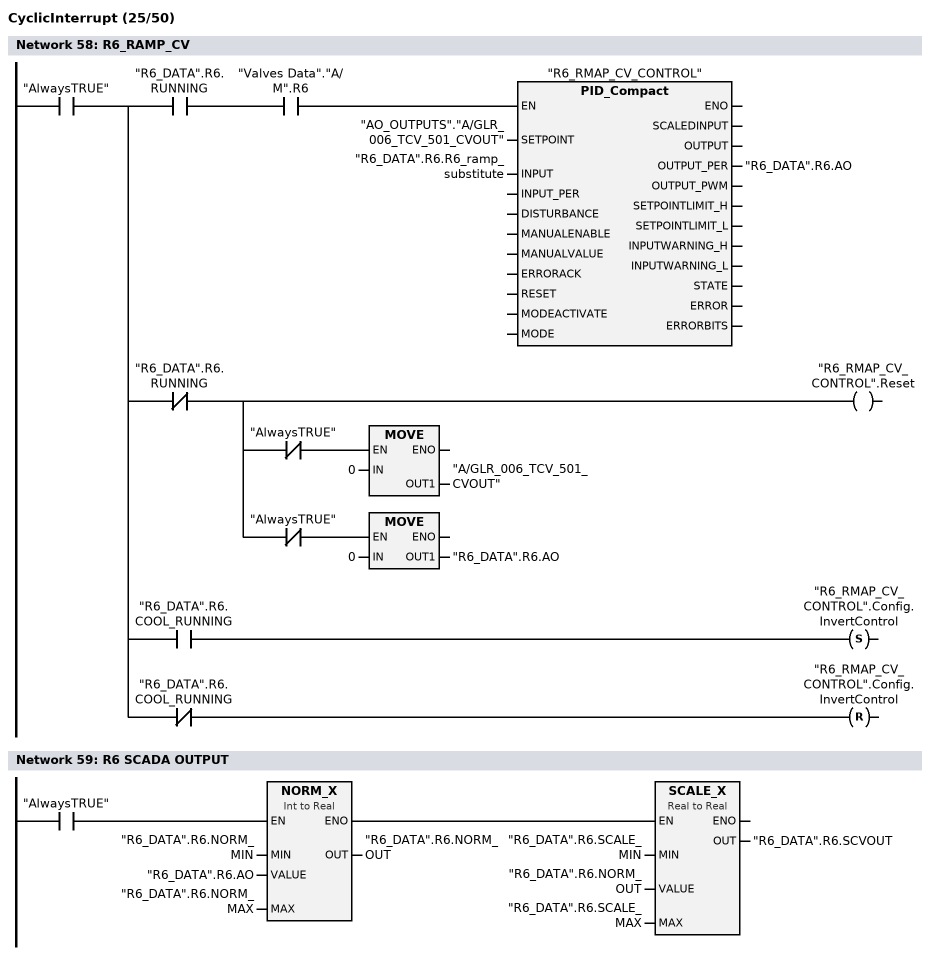
   RUNG wire#powerrail
      Contact( "AlwaysTRUE" )
      wire#w1
      Contact( "R6_DATA".R6.RUNNING )
      Contact( "Valves Data"."A/M".R6 )
      "R6_RMAP_CV_CONTROL".PID_Compact(Setpoint := "AO_OUTPUTS"."A/GLR_006_TCV_501_CVOUT", Input := "R6_DATA".R6.R6_ramp_substitute, Input_PER :=, Disturbance :=, ManualEnable :=, ManualValue :=, ErrorAck :=, Reset :=, ModeActivate :=, Mode :=, ScaledInput =>, Output =>, Output_PER => "R6_DATA".R6.AO, Output_PWM =>, SetpointLimit_H =>, SetpointLimit_L =>, InputWarning_H =>, InputWarning_L =>, State =>, Error =>, ErrorBits =>)
   END_RUNG
   RUNG wire#w1
      I_Contact( "R6_DATA".R6.RUNNING )
      wire#w2
      Coil( "R6_RMAP_CV_CONTROL".Reset )
   END_RUNG
   RUNG wire#w2
      I_Contact( "AlwaysTRUE" )
      Move(in := 0, out1 => "A/GLR_006_TCV_501_CVOUT")
   END_RUNG
   RUNG wire#w2
      I_Contact( "AlwaysTRUE" )
      Move(in := 0, out1 => "R6_DATA".R6.AO)
   END_RUNG
   RUNG wire#w1
      Contact( "R6_DATA".R6.COOL_RUNNING )
      S_Coil( "R6_RMAP_CV_CONTROL".Config.InvertControl )
   END_RUNG
   RUNG wire#w1
      I_Contact( "R6_DATA".R6.COOL_RUNNING )
      R_Coil( "R6_RMAP_CV_CONTROL".Config.InvertControl )
   END_RUNG
   // the same network as SCL:
   #_w1 := "AlwaysTRUE";
   IF "AlwaysTRUE" AND "R6_DATA".R6.RUNNING AND "Valves Data"."A/M".R6 THEN
       "R6_RMAP_CV_CONTROL"(Setpoint := "AO_OUTPUTS"."A/GLR_006_TCV_501_CVOUT",   // PID_Compact
                            Input := "R6_DATA".R6.R6_ramp_substitute,
                            Output_PER => "R6_DATA".R6.AO);
   END_IF;
   "R6_RMAP_CV_CONTROL".Reset := #_w1 AND NOT "R6_DATA".R6.RUNNING;
   IF "R6_RMAP_CV_CONTROL".Reset AND NOT "AlwaysTRUE" THEN
       "A/GLR_006_TCV_501_CVOUT" := 0;
       "R6_DATA".R6.AO := 0;
   END_IF;
   IF #_w1 AND "R6_DATA".R6.COOL_RUNNING THEN "R6_RMAP_CV_CONTROL".Config.InvertControl := TRUE; END_IF;
   IF #_w1 AND NOT "R6_DATA".R6.COOL_RUNNING THEN "R6_RMAP_CV_CONTROL".Config.InvertControl := FALSE; END_IF;
END_REGION

REGION Network 59: R6 SCADA OUTPUT
   RUNG wire#powerrail
      Contact( "AlwaysTRUE" )
      { S7_Templates := "[SrcType := Int, DestType := Real]" } Normalize(min := "R6_DATA".R6.NORM_MIN, value := "R6_DATA".R6.AO, max := "R6_DATA".R6.NORM_MAX, out => "R6_DATA".R6.NORM_OUT)
      { S7_Templates := "[SrcType := Real, DestType := Real]" } Scale(min := "R6_DATA".R6.SCALE_MIN, value := "R6_DATA".R6.NORM_OUT, max := "R6_DATA".R6.SCALE_MAX, out => "R6_DATA".R6.SCVOUT)
   END_RUNG
   // the same network as SCL:
   IF "AlwaysTRUE" THEN
       "R6_DATA".R6.NORM_OUT := NORM_X(MIN := "R6_DATA".R6.NORM_MIN, VALUE := "R6_DATA".R6.AO, MAX := "R6_DATA".R6.NORM_MAX);
       "R6_DATA".R6.SCVOUT := SCALE_X(MIN := "R6_DATA".R6.SCALE_MIN, VALUE := "R6_DATA".R6.NORM_OUT, MAX := "R6_DATA".R6.SCALE_MAX);
   END_IF;
END_REGION

REGION Network 60: R6 AUTO/MANUAL OUTPUT
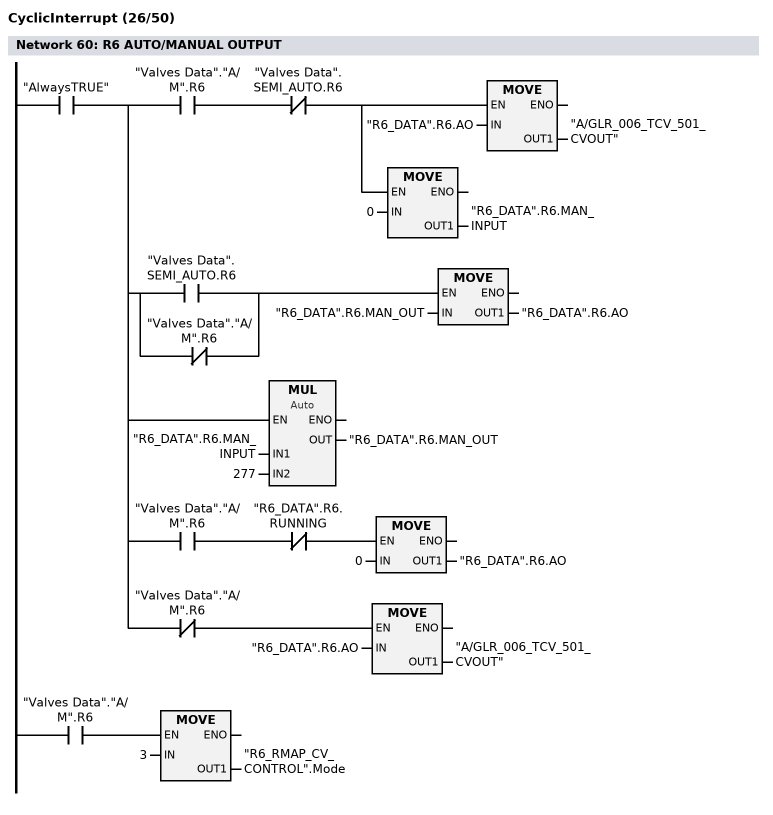
   RUNG wire#powerrail
      Contact( "AlwaysTRUE" )
      wire#w1
      Contact( "Valves Data"."A/M".R6 )
      I_Contact( "Valves Data".SEMI_AUTO.R6 )
      wire#w2
      Move(in := "R6_DATA".R6.AO, out1 => "A/GLR_006_TCV_501_CVOUT")
   END_RUNG
   RUNG wire#w2
      Move(in := 0, out1 => "R6_DATA".R6.MAN_INPUT)
   END_RUNG
   RUNG wire#w1
      Contact( "Valves Data".SEMI_AUTO.R6 )
      wire#w3
      Move(in := "R6_DATA".R6.MAN_OUT, out1 => "R6_DATA".R6.AO)
   END_RUNG
   RUNG wire#w1
      I_Contact( "Valves Data"."A/M".R6 )
   END_RUNG wire#w3
   RUNG wire#w1
      Mul(in1 := "R6_DATA".R6.MAN_INPUT, in2 := 277, out => "R6_DATA".R6.MAN_OUT)
   END_RUNG
   RUNG wire#w1
      Contact( "Valves Data"."A/M".R6 )
      I_Contact( "R6_DATA".R6.RUNNING )
      Move(in := 0, out1 => "R6_DATA".R6.AO)
   END_RUNG
   RUNG wire#w1
      I_Contact( "Valves Data"."A/M".R6 )
      Move(in := "R6_DATA".R6.AO, out1 => "A/GLR_006_TCV_501_CVOUT")
   END_RUNG
   RUNG wire#powerrail
      Contact( "Valves Data"."A/M".R6 )
      Move(in := 3, out1 => "R6_RMAP_CV_CONTROL".Mode)
   END_RUNG
   // the same network as SCL:
   IF "AlwaysTRUE" AND "Valves Data"."A/M".R6 AND NOT "Valves Data".SEMI_AUTO.R6 THEN
       "A/GLR_006_TCV_501_CVOUT" := "R6_DATA".R6.AO;
       "R6_DATA".R6.MAN_INPUT := 0;
   END_IF;
   IF "AlwaysTRUE" AND ("Valves Data".SEMI_AUTO.R6 OR NOT "Valves Data"."A/M".R6) THEN
       "R6_DATA".R6.AO := "R6_DATA".R6.MAN_OUT;
   END_IF;
   IF "AlwaysTRUE" THEN "R6_DATA".R6.MAN_OUT := "R6_DATA".R6.MAN_INPUT * 277; END_IF;
   IF "AlwaysTRUE" AND "Valves Data"."A/M".R6 AND NOT "R6_DATA".R6.RUNNING THEN "R6_DATA".R6.AO := 0; END_IF;
   IF "AlwaysTRUE" AND NOT "Valves Data"."A/M".R6 THEN "A/GLR_006_TCV_501_CVOUT" := "R6_DATA".R6.AO; END_IF;
   IF "Valves Data"."A/M".R6 THEN "R6_RMAP_CV_CONTROL".Mode := 3; END_IF;
END_REGION

REGION Network 61: R7_RAMP_CV
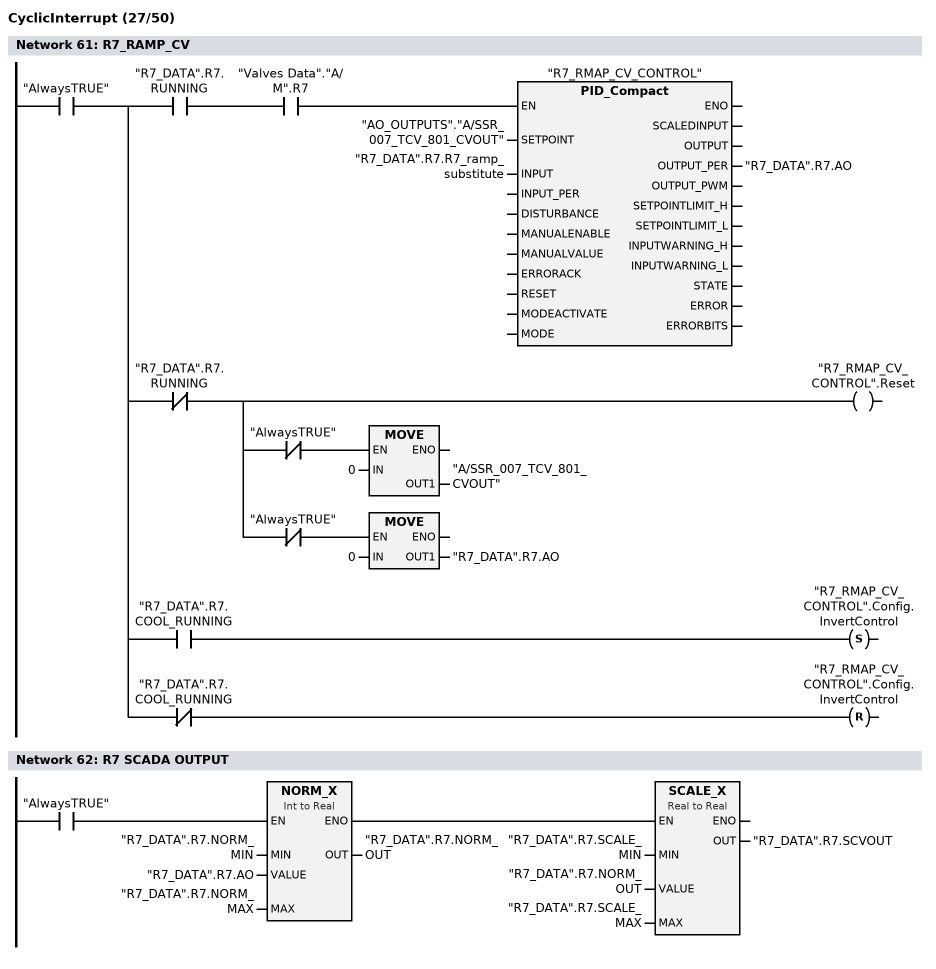
   RUNG wire#powerrail
      Contact( "AlwaysTRUE" )
      wire#w1
      Contact( "R7_DATA".R7.RUNNING )
      Contact( "Valves Data"."A/M".R7 )
      "R7_RMAP_CV_CONTROL".PID_Compact(Setpoint := "AO_OUTPUTS"."A/SSR_007_TCV_801_CVOUT", Input := "R7_DATA".R7.R7_ramp_substitute, Input_PER :=, Disturbance :=, ManualEnable :=, ManualValue :=, ErrorAck :=, Reset :=, ModeActivate :=, Mode :=, ScaledInput =>, Output =>, Output_PER => "R7_DATA".R7.AO, Output_PWM =>, SetpointLimit_H =>, SetpointLimit_L =>, InputWarning_H =>, InputWarning_L =>, State =>, Error =>, ErrorBits =>)
   END_RUNG
   RUNG wire#w1
      I_Contact( "R7_DATA".R7.RUNNING )
      wire#w2
      Coil( "R7_RMAP_CV_CONTROL".Reset )
   END_RUNG
   RUNG wire#w2
      I_Contact( "AlwaysTRUE" )
      Move(in := 0, out1 => "A/SSR_007_TCV_801_CVOUT")
   END_RUNG
   RUNG wire#w2
      I_Contact( "AlwaysTRUE" )
      Move(in := 0, out1 => "R7_DATA".R7.AO)
   END_RUNG
   RUNG wire#w1
      Contact( "R7_DATA".R7.COOL_RUNNING )
      S_Coil( "R7_RMAP_CV_CONTROL".Config.InvertControl )
   END_RUNG
   RUNG wire#w1
      I_Contact( "R7_DATA".R7.COOL_RUNNING )
      R_Coil( "R7_RMAP_CV_CONTROL".Config.InvertControl )
   END_RUNG
   // the same network as SCL:
   #_w1 := "AlwaysTRUE";
   IF "AlwaysTRUE" AND "R7_DATA".R7.RUNNING AND "Valves Data"."A/M".R7 THEN
       "R7_RMAP_CV_CONTROL"(Setpoint := "AO_OUTPUTS"."A/SSR_007_TCV_801_CVOUT",   // PID_Compact
                            Input := "R7_DATA".R7.R7_ramp_substitute,
                            Output_PER => "R7_DATA".R7.AO);
   END_IF;
   "R7_RMAP_CV_CONTROL".Reset := #_w1 AND NOT "R7_DATA".R7.RUNNING;
   IF "R7_RMAP_CV_CONTROL".Reset AND NOT "AlwaysTRUE" THEN
       "A/SSR_007_TCV_801_CVOUT" := 0;
       "R7_DATA".R7.AO := 0;
   END_IF;
   IF #_w1 AND "R7_DATA".R7.COOL_RUNNING THEN "R7_RMAP_CV_CONTROL".Config.InvertControl := TRUE; END_IF;
   IF #_w1 AND NOT "R7_DATA".R7.COOL_RUNNING THEN "R7_RMAP_CV_CONTROL".Config.InvertControl := FALSE; END_IF;
END_REGION

REGION Network 62: R7 SCADA OUTPUT
   RUNG wire#powerrail
      Contact( "AlwaysTRUE" )
      { S7_Templates := "[SrcType := Int, DestType := Real]" } Normalize(min := "R7_DATA".R7.NORM_MIN, value := "R7_DATA".R7.AO, max := "R7_DATA".R7.NORM_MAX, out => "R7_DATA".R7.NORM_OUT)
      { S7_Templates := "[SrcType := Real, DestType := Real]" } Scale(min := "R7_DATA".R7.SCALE_MIN, value := "R7_DATA".R7.NORM_OUT, max := "R7_DATA".R7.SCALE_MAX, out => "R7_DATA".R7.SCVOUT)
   END_RUNG
   // the same network as SCL:
   IF "AlwaysTRUE" THEN
       "R7_DATA".R7.NORM_OUT := NORM_X(MIN := "R7_DATA".R7.NORM_MIN, VALUE := "R7_DATA".R7.AO, MAX := "R7_DATA".R7.NORM_MAX);
       "R7_DATA".R7.SCVOUT := SCALE_X(MIN := "R7_DATA".R7.SCALE_MIN, VALUE := "R7_DATA".R7.NORM_OUT, MAX := "R7_DATA".R7.SCALE_MAX);
   END_IF;
END_REGION

REGION Network 63: R7 AUTO/MANUAL OUTPUT
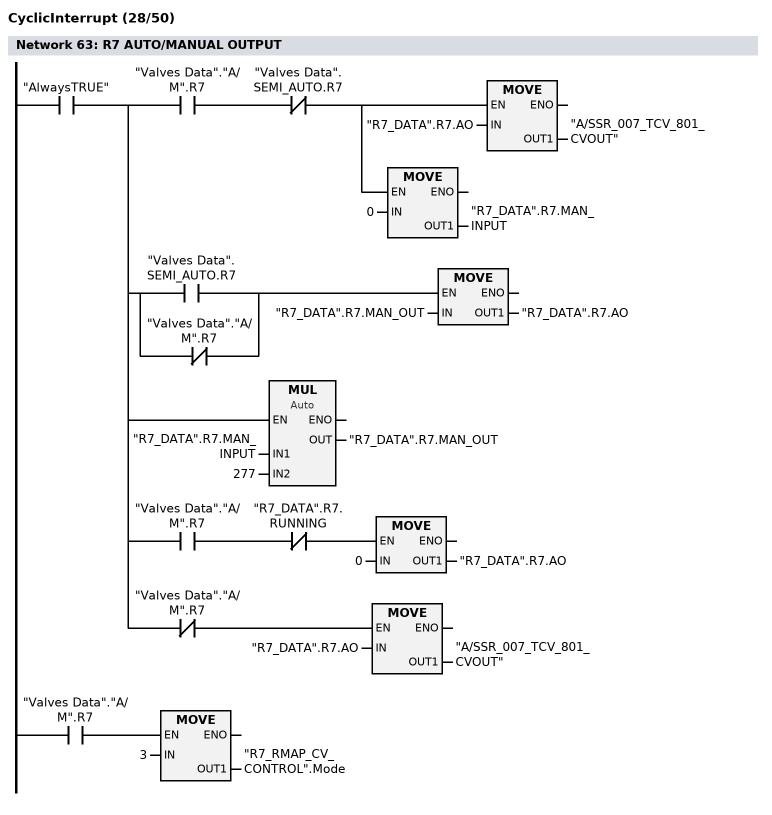
   RUNG wire#powerrail
      Contact( "AlwaysTRUE" )
      wire#w1
      Contact( "Valves Data"."A/M".R7 )
      I_Contact( "Valves Data".SEMI_AUTO.R7 )
      wire#w2
      Move(in := "R7_DATA".R7.AO, out1 => "A/SSR_007_TCV_801_CVOUT")
   END_RUNG
   RUNG wire#w2
      Move(in := 0, out1 => "R7_DATA".R7.MAN_INPUT)
   END_RUNG
   RUNG wire#w1
      Contact( "Valves Data".SEMI_AUTO.R7 )
      wire#w3
      Move(in := "R7_DATA".R7.MAN_OUT, out1 => "R7_DATA".R7.AO)
   END_RUNG
   RUNG wire#w1
      I_Contact( "Valves Data"."A/M".R7 )
   END_RUNG wire#w3
   RUNG wire#w1
      Mul(in1 := "R7_DATA".R7.MAN_INPUT, in2 := 277, out => "R7_DATA".R7.MAN_OUT)
   END_RUNG
   RUNG wire#w1
      Contact( "Valves Data"."A/M".R7 )
      I_Contact( "R7_DATA".R7.RUNNING )
      Move(in := 0, out1 => "R7_DATA".R7.AO)
   END_RUNG
   RUNG wire#w1
      I_Contact( "Valves Data"."A/M".R7 )
      Move(in := "R7_DATA".R7.AO, out1 => "A/SSR_007_TCV_801_CVOUT")
   END_RUNG
   RUNG wire#powerrail
      Contact( "Valves Data"."A/M".R7 )
      Move(in := 3, out1 => "R7_RMAP_CV_CONTROL".Mode)
   END_RUNG
   // the same network as SCL:
   IF "AlwaysTRUE" AND "Valves Data"."A/M".R7 AND NOT "Valves Data".SEMI_AUTO.R7 THEN
       "A/SSR_007_TCV_801_CVOUT" := "R7_DATA".R7.AO;
       "R7_DATA".R7.MAN_INPUT := 0;
   END_IF;
   IF "AlwaysTRUE" AND ("Valves Data".SEMI_AUTO.R7 OR NOT "Valves Data"."A/M".R7) THEN
       "R7_DATA".R7.AO := "R7_DATA".R7.MAN_OUT;
   END_IF;
   IF "AlwaysTRUE" THEN "R7_DATA".R7.MAN_OUT := "R7_DATA".R7.MAN_INPUT * 277; END_IF;
   IF "AlwaysTRUE" AND "Valves Data"."A/M".R7 AND NOT "R7_DATA".R7.RUNNING THEN "R7_DATA".R7.AO := 0; END_IF;
   IF "AlwaysTRUE" AND NOT "Valves Data"."A/M".R7 THEN "A/SSR_007_TCV_801_CVOUT" := "R7_DATA".R7.AO; END_IF;
   IF "Valves Data"."A/M".R7 THEN "R7_RMAP_CV_CONTROL".Mode := 3; END_IF;
END_REGION

REGION Network 64: R8_RAMP_CV
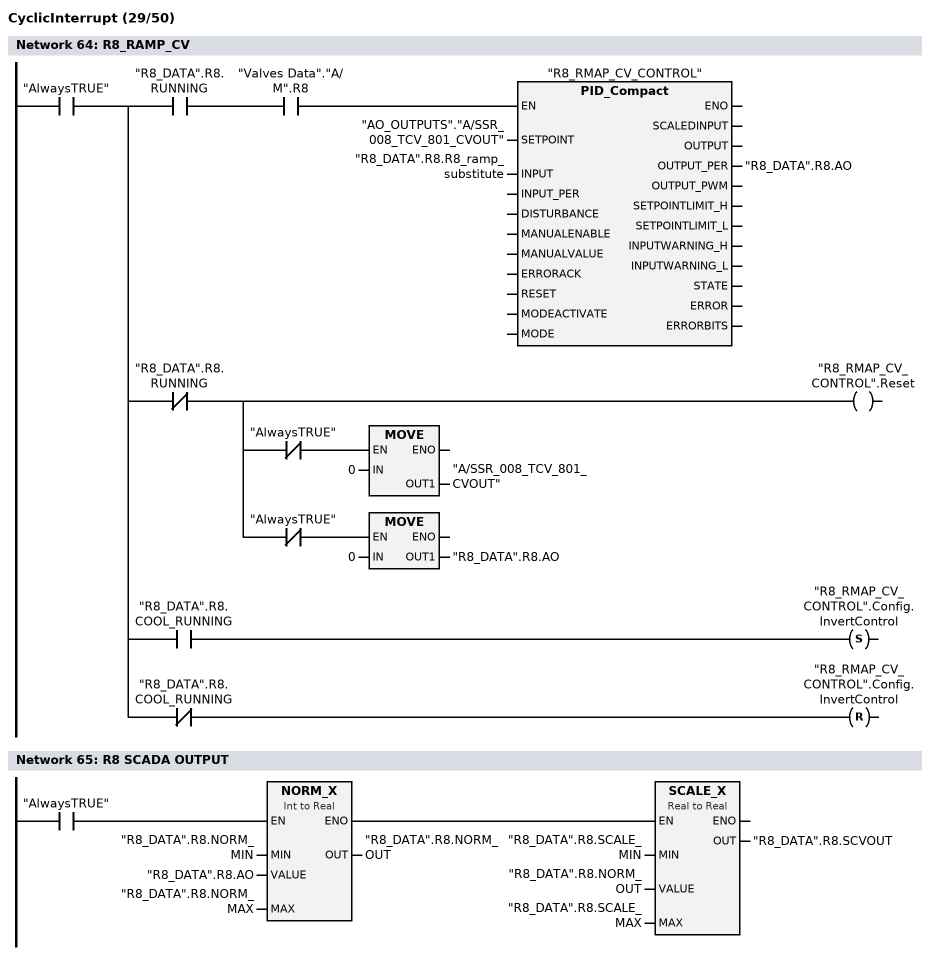
   RUNG wire#powerrail
      Contact( "AlwaysTRUE" )
      wire#w1
      Contact( "R8_DATA".R8.RUNNING )
      Contact( "Valves Data"."A/M".R8 )
      "R8_RMAP_CV_CONTROL".PID_Compact(Setpoint := "AO_OUTPUTS"."A/SSR_008_TCV_801_CVOUT", Input := "R8_DATA".R8.R8_ramp_substitute, Input_PER :=, Disturbance :=, ManualEnable :=, ManualValue :=, ErrorAck :=, Reset :=, ModeActivate :=, Mode :=, ScaledInput =>, Output =>, Output_PER => "R8_DATA".R8.AO, Output_PWM =>, SetpointLimit_H =>, SetpointLimit_L =>, InputWarning_H =>, InputWarning_L =>, State =>, Error =>, ErrorBits =>)
   END_RUNG
   RUNG wire#w1
      I_Contact( "R8_DATA".R8.RUNNING )
      wire#w2
      Coil( "R8_RMAP_CV_CONTROL".Reset )
   END_RUNG
   RUNG wire#w2
      I_Contact( "AlwaysTRUE" )
      Move(in := 0, out1 => "A/SSR_008_TCV_801_CVOUT")
   END_RUNG
   RUNG wire#w2
      I_Contact( "AlwaysTRUE" )
      Move(in := 0, out1 => "R8_DATA".R8.AO)
   END_RUNG
   RUNG wire#w1
      Contact( "R8_DATA".R8.COOL_RUNNING )
      S_Coil( "R8_RMAP_CV_CONTROL".Config.InvertControl )
   END_RUNG
   RUNG wire#w1
      I_Contact( "R8_DATA".R8.COOL_RUNNING )
      R_Coil( "R8_RMAP_CV_CONTROL".Config.InvertControl )
   END_RUNG
   // the same network as SCL:
   #_w1 := "AlwaysTRUE";
   IF "AlwaysTRUE" AND "R8_DATA".R8.RUNNING AND "Valves Data"."A/M".R8 THEN
       "R8_RMAP_CV_CONTROL"(Setpoint := "AO_OUTPUTS"."A/SSR_008_TCV_801_CVOUT",   // PID_Compact
                            Input := "R8_DATA".R8.R8_ramp_substitute,
                            Output_PER => "R8_DATA".R8.AO);
   END_IF;
   "R8_RMAP_CV_CONTROL".Reset := #_w1 AND NOT "R8_DATA".R8.RUNNING;
   IF "R8_RMAP_CV_CONTROL".Reset AND NOT "AlwaysTRUE" THEN
       "A/SSR_008_TCV_801_CVOUT" := 0;
       "R8_DATA".R8.AO := 0;
   END_IF;
   IF #_w1 AND "R8_DATA".R8.COOL_RUNNING THEN "R8_RMAP_CV_CONTROL".Config.InvertControl := TRUE; END_IF;
   IF #_w1 AND NOT "R8_DATA".R8.COOL_RUNNING THEN "R8_RMAP_CV_CONTROL".Config.InvertControl := FALSE; END_IF;
END_REGION

REGION Network 65: R8 SCADA OUTPUT
   RUNG wire#powerrail
      Contact( "AlwaysTRUE" )
      { S7_Templates := "[SrcType := Int, DestType := Real]" } Normalize(min := "R8_DATA".R8.NORM_MIN, value := "R8_DATA".R8.AO, max := "R8_DATA".R8.NORM_MAX, out => "R8_DATA".R8.NORM_OUT)
      { S7_Templates := "[SrcType := Real, DestType := Real]" } Scale(min := "R8_DATA".R8.SCALE_MIN, value := "R8_DATA".R8.NORM_OUT, max := "R8_DATA".R8.SCALE_MAX, out => "R8_DATA".R8.SCVOUT)
   END_RUNG
   // the same network as SCL:
   IF "AlwaysTRUE" THEN
       "R8_DATA".R8.NORM_OUT := NORM_X(MIN := "R8_DATA".R8.NORM_MIN, VALUE := "R8_DATA".R8.AO, MAX := "R8_DATA".R8.NORM_MAX);
       "R8_DATA".R8.SCVOUT := SCALE_X(MIN := "R8_DATA".R8.SCALE_MIN, VALUE := "R8_DATA".R8.NORM_OUT, MAX := "R8_DATA".R8.SCALE_MAX);
   END_IF;
END_REGION

REGION Network 66: R8 AUTO/MANUAL OUTPUT
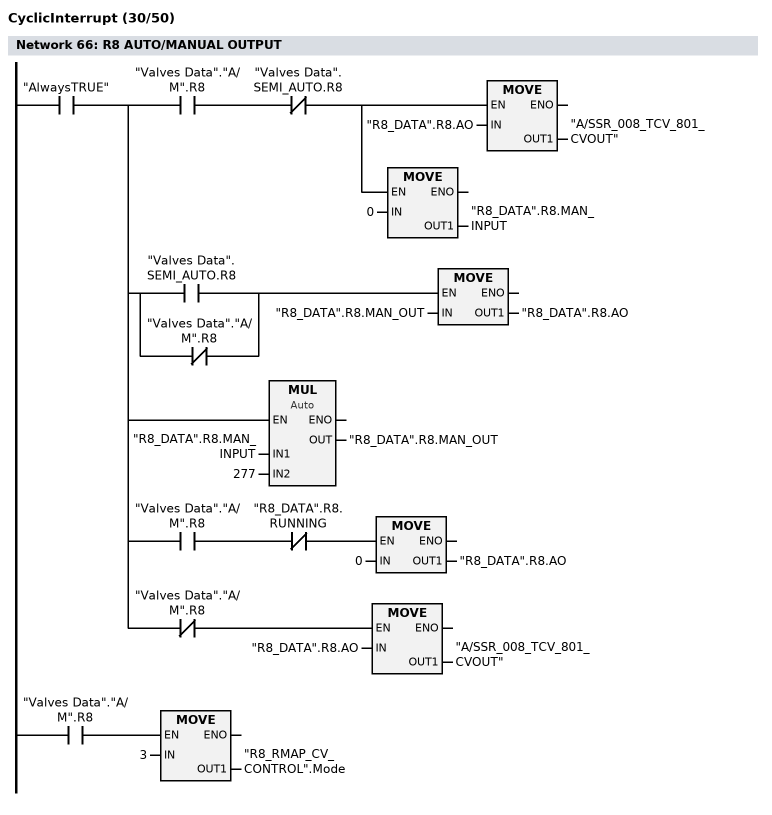
   RUNG wire#powerrail
      Contact( "AlwaysTRUE" )
      wire#w1
      Contact( "Valves Data"."A/M".R8 )
      I_Contact( "Valves Data".SEMI_AUTO.R8 )
      wire#w2
      Move(in := "R8_DATA".R8.AO, out1 => "A/SSR_008_TCV_801_CVOUT")
   END_RUNG
   RUNG wire#w2
      Move(in := 0, out1 => "R8_DATA".R8.MAN_INPUT)
   END_RUNG
   RUNG wire#w1
      Contact( "Valves Data".SEMI_AUTO.R8 )
      wire#w3
      Move(in := "R8_DATA".R8.MAN_OUT, out1 => "R8_DATA".R8.AO)
   END_RUNG
   RUNG wire#w1
      I_Contact( "Valves Data"."A/M".R8 )
   END_RUNG wire#w3
   RUNG wire#w1
      Mul(in1 := "R8_DATA".R8.MAN_INPUT, in2 := 277, out => "R8_DATA".R8.MAN_OUT)
   END_RUNG
   RUNG wire#w1
      Contact( "Valves Data"."A/M".R8 )
      I_Contact( "R8_DATA".R8.RUNNING )
      Move(in := 0, out1 => "R8_DATA".R8.AO)
   END_RUNG
   RUNG wire#w1
      I_Contact( "Valves Data"."A/M".R8 )
      Move(in := "R8_DATA".R8.AO, out1 => "A/SSR_008_TCV_801_CVOUT")
   END_RUNG
   RUNG wire#powerrail
      Contact( "Valves Data"."A/M".R8 )
      Move(in := 3, out1 => "R8_RMAP_CV_CONTROL".Mode)
   END_RUNG
   // the same network as SCL:
   IF "AlwaysTRUE" AND "Valves Data"."A/M".R8 AND NOT "Valves Data".SEMI_AUTO.R8 THEN
       "A/SSR_008_TCV_801_CVOUT" := "R8_DATA".R8.AO;
       "R8_DATA".R8.MAN_INPUT := 0;
   END_IF;
   IF "AlwaysTRUE" AND ("Valves Data".SEMI_AUTO.R8 OR NOT "Valves Data"."A/M".R8) THEN
       "R8_DATA".R8.AO := "R8_DATA".R8.MAN_OUT;
   END_IF;
   IF "AlwaysTRUE" THEN "R8_DATA".R8.MAN_OUT := "R8_DATA".R8.MAN_INPUT * 277; END_IF;
   IF "AlwaysTRUE" AND "Valves Data"."A/M".R8 AND NOT "R8_DATA".R8.RUNNING THEN "R8_DATA".R8.AO := 0; END_IF;
   IF "AlwaysTRUE" AND NOT "Valves Data"."A/M".R8 THEN "A/SSR_008_TCV_801_CVOUT" := "R8_DATA".R8.AO; END_IF;
   IF "Valves Data"."A/M".R8 THEN "R8_RMAP_CV_CONTROL".Mode := 3; END_IF;
END_REGION

REGION Network 67: R9_RAMP_CV
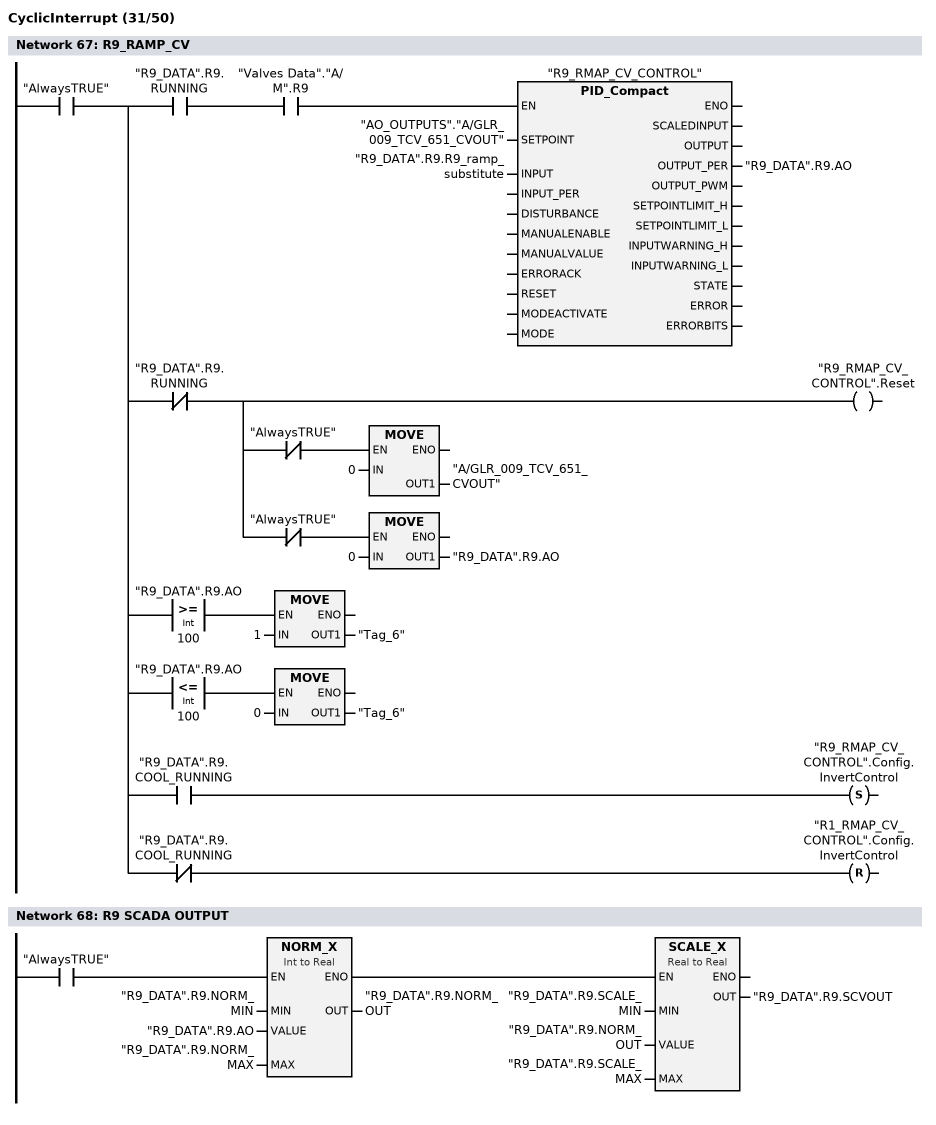
   RUNG wire#powerrail
      Contact( "AlwaysTRUE" )
      wire#w1
      Contact( "R9_DATA".R9.RUNNING )
      Contact( "Valves Data"."A/M".R9 )
      "R9_RMAP_CV_CONTROL".PID_Compact(Setpoint := "AO_OUTPUTS"."A/GLR_009_TCV_651_CVOUT", Input := "R9_DATA".R9.R9_ramp_substitute, Input_PER :=, Disturbance :=, ManualEnable :=, ManualValue :=, ErrorAck :=, Reset :=, ModeActivate :=, Mode :=, ScaledInput =>, Output =>, Output_PER => "R9_DATA".R9.AO, Output_PWM =>, SetpointLimit_H =>, SetpointLimit_L =>, InputWarning_H =>, InputWarning_L =>, State =>, Error =>, ErrorBits =>)
   END_RUNG
   RUNG wire#w1
      I_Contact( "R9_DATA".R9.RUNNING )
      wire#w2
      Coil( "R9_RMAP_CV_CONTROL".Reset )
   END_RUNG
   RUNG wire#w2
      I_Contact( "AlwaysTRUE" )
      Move(in := 0, out1 => "A/GLR_009_TCV_651_CVOUT")
   END_RUNG
   RUNG wire#w2
      I_Contact( "AlwaysTRUE" )
      Move(in := 0, out1 => "R9_DATA".R9.AO)
   END_RUNG
   RUNG wire#w1
      { S7_Templates := "SrcType := Int" } GE_Contact(in1 := "R9_DATA".R9.AO, in2 := 100)
      Move(in := 1, out1 => "Tag_6")
   END_RUNG
   RUNG wire#w1
      { S7_Templates := "SrcType := Int" } LE_Contact(in1 := "R9_DATA".R9.AO, in2 := 100)
      Move(in := 0, out1 => "Tag_6")
   END_RUNG
   RUNG wire#w1
      Contact( "R9_DATA".R9.COOL_RUNNING )
      S_Coil( "R9_RMAP_CV_CONTROL".Config.InvertControl )
   END_RUNG
   RUNG wire#w1
      I_Contact( "R9_DATA".R9.COOL_RUNNING )
      R_Coil( "R1_RMAP_CV_CONTROL".Config.InvertControl )
   END_RUNG
   // the same network as SCL:
   #_w1 := "AlwaysTRUE";
   IF "AlwaysTRUE" AND "R9_DATA".R9.RUNNING AND "Valves Data"."A/M".R9 THEN
       "R9_RMAP_CV_CONTROL"(Setpoint := "AO_OUTPUTS"."A/GLR_009_TCV_651_CVOUT",   // PID_Compact
                            Input := "R9_DATA".R9.R9_ramp_substitute,
                            Output_PER => "R9_DATA".R9.AO);
   END_IF;
   "R9_RMAP_CV_CONTROL".Reset := #_w1 AND NOT "R9_DATA".R9.RUNNING;
   IF "R9_RMAP_CV_CONTROL".Reset AND NOT "AlwaysTRUE" THEN
       "A/GLR_009_TCV_651_CVOUT" := 0;
       "R9_DATA".R9.AO := 0;
   END_IF;
   IF #_w1 AND ("R9_DATA".R9.AO >= 100) THEN "Tag_6" := 1; END_IF;
   IF #_w1 AND ("R9_DATA".R9.AO <= 100) THEN "Tag_6" := 0; END_IF;
   IF #_w1 AND "R9_DATA".R9.COOL_RUNNING THEN "R9_RMAP_CV_CONTROL".Config.InvertControl := TRUE; END_IF;
   IF #_w1 AND NOT "R9_DATA".R9.COOL_RUNNING THEN "R1_RMAP_CV_CONTROL".Config.InvertControl := FALSE; END_IF;
END_REGION

REGION Network 68: R9 SCADA OUTPUT
   RUNG wire#powerrail
      Contact( "AlwaysTRUE" )
      { S7_Templates := "[SrcType := Int, DestType := Real]" } Normalize(min := "R9_DATA".R9.NORM_MIN, value := "R9_DATA".R9.AO, max := "R9_DATA".R9.NORM_MAX, out => "R9_DATA".R9.NORM_OUT)
      { S7_Templates := "[SrcType := Real, DestType := Real]" } Scale(min := "R9_DATA".R9.SCALE_MIN, value := "R9_DATA".R9.NORM_OUT, max := "R9_DATA".R9.SCALE_MAX, out => "R9_DATA".R9.SCVOUT)
   END_RUNG
   // the same network as SCL:
   IF "AlwaysTRUE" THEN
       "R9_DATA".R9.NORM_OUT := NORM_X(MIN := "R9_DATA".R9.NORM_MIN, VALUE := "R9_DATA".R9.AO, MAX := "R9_DATA".R9.NORM_MAX);
       "R9_DATA".R9.SCVOUT := SCALE_X(MIN := "R9_DATA".R9.SCALE_MIN, VALUE := "R9_DATA".R9.NORM_OUT, MAX := "R9_DATA".R9.SCALE_MAX);
   END_IF;
END_REGION

REGION Network 69: R9 AUTO/MANUAL OUTPUT
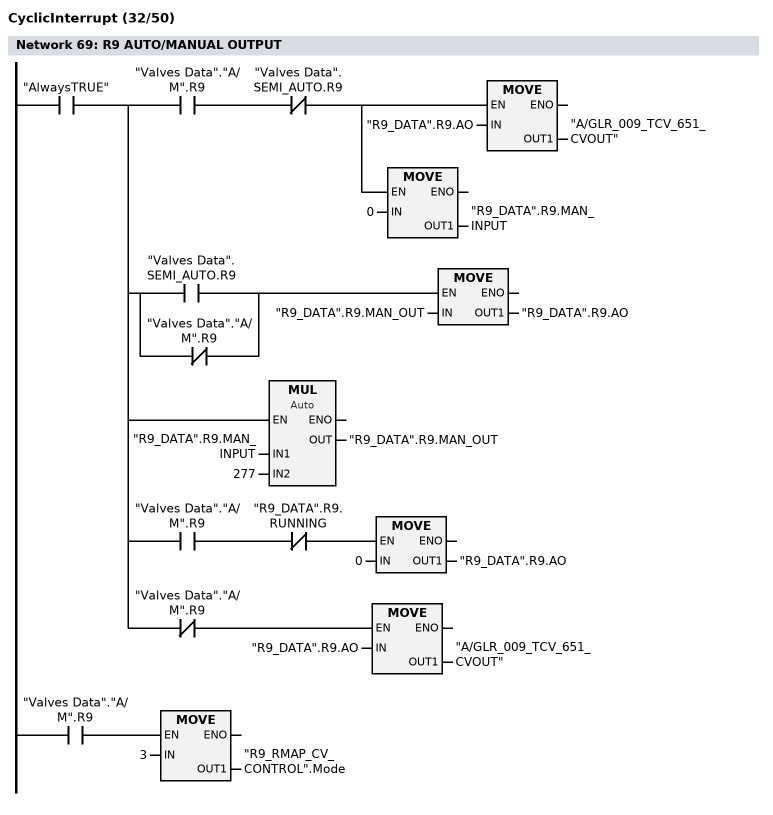
   RUNG wire#powerrail
      Contact( "AlwaysTRUE" )
      wire#w1
      Contact( "Valves Data"."A/M".R9 )
      I_Contact( "Valves Data".SEMI_AUTO.R9 )
      wire#w2
      Move(in := "R9_DATA".R9.AO, out1 => "A/GLR_009_TCV_651_CVOUT")
   END_RUNG
   RUNG wire#w2
      Move(in := 0, out1 => "R9_DATA".R9.MAN_INPUT)
   END_RUNG
   RUNG wire#w1
      Contact( "Valves Data".SEMI_AUTO.R9 )
      wire#w3
      Move(in := "R9_DATA".R9.MAN_OUT, out1 => "R9_DATA".R9.AO)
   END_RUNG
   RUNG wire#w1
      I_Contact( "Valves Data"."A/M".R9 )
   END_RUNG wire#w3
   RUNG wire#w1
      Mul(in1 := "R9_DATA".R9.MAN_INPUT, in2 := 277, out => "R9_DATA".R9.MAN_OUT)
   END_RUNG
   RUNG wire#w1
      Contact( "Valves Data"."A/M".R9 )
      I_Contact( "R9_DATA".R9.RUNNING )
      Move(in := 0, out1 => "R9_DATA".R9.AO)
   END_RUNG
   RUNG wire#w1
      I_Contact( "Valves Data"."A/M".R9 )
      Move(in := "R9_DATA".R9.AO, out1 => "A/GLR_009_TCV_651_CVOUT")
   END_RUNG
   RUNG wire#powerrail
      Contact( "Valves Data"."A/M".R9 )
      Move(in := 3, out1 => "R9_RMAP_CV_CONTROL".Mode)
   END_RUNG
   // the same network as SCL:
   IF "AlwaysTRUE" AND "Valves Data"."A/M".R9 AND NOT "Valves Data".SEMI_AUTO.R9 THEN
       "A/GLR_009_TCV_651_CVOUT" := "R9_DATA".R9.AO;
       "R9_DATA".R9.MAN_INPUT := 0;
   END_IF;
   IF "AlwaysTRUE" AND ("Valves Data".SEMI_AUTO.R9 OR NOT "Valves Data"."A/M".R9) THEN
       "R9_DATA".R9.AO := "R9_DATA".R9.MAN_OUT;
   END_IF;
   IF "AlwaysTRUE" THEN "R9_DATA".R9.MAN_OUT := "R9_DATA".R9.MAN_INPUT * 277; END_IF;
   IF "AlwaysTRUE" AND "Valves Data"."A/M".R9 AND NOT "R9_DATA".R9.RUNNING THEN "R9_DATA".R9.AO := 0; END_IF;
   IF "AlwaysTRUE" AND NOT "Valves Data"."A/M".R9 THEN "A/GLR_009_TCV_651_CVOUT" := "R9_DATA".R9.AO; END_IF;
   IF "Valves Data"."A/M".R9 THEN "R9_RMAP_CV_CONTROL".Mode := 3; END_IF;
END_REGION

REGION Network 70: R10_RAMP_CV
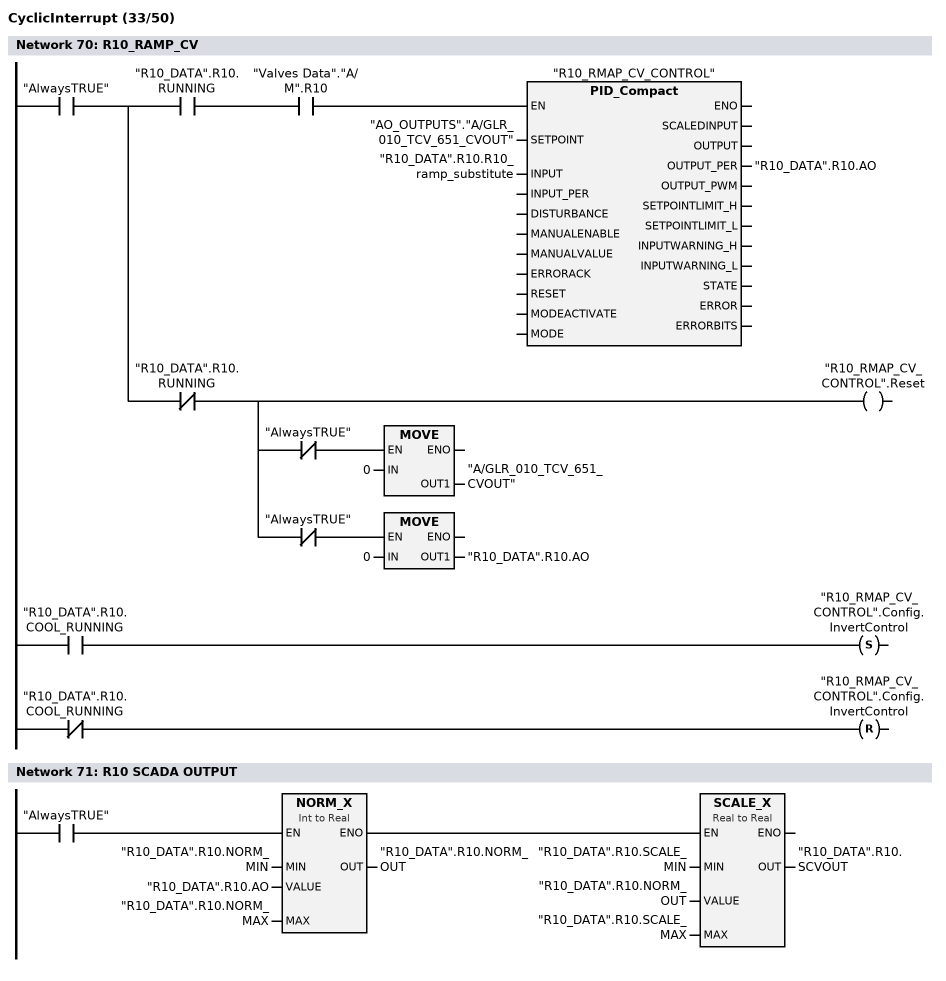
   RUNG wire#powerrail
      Contact( "AlwaysTRUE" )
      wire#w1
      Contact( "R10_DATA".R10.RUNNING )
      Contact( "Valves Data"."A/M".R10 )
      "R10_RMAP_CV_CONTROL".PID_Compact(Setpoint := "AO_OUTPUTS"."A/GLR_010_TCV_651_CVOUT", Input := "R10_DATA".R10.R10_ramp_substitute, Input_PER :=, Disturbance :=, ManualEnable :=, ManualValue :=, ErrorAck :=, Reset :=, ModeActivate :=, Mode :=, ScaledInput =>, Output =>, Output_PER => "R10_DATA".R10.AO, Output_PWM =>, SetpointLimit_H =>, SetpointLimit_L =>, InputWarning_H =>, InputWarning_L =>, State =>, Error =>, ErrorBits =>)
   END_RUNG
   RUNG wire#w1
      I_Contact( "R10_DATA".R10.RUNNING )
      wire#w2
      Coil( "R10_RMAP_CV_CONTROL".Reset )
   END_RUNG
   RUNG wire#w2
      I_Contact( "AlwaysTRUE" )
      Move(in := 0, out1 => "A/GLR_010_TCV_651_CVOUT")
   END_RUNG
   RUNG wire#w2
      I_Contact( "AlwaysTRUE" )
      Move(in := 0, out1 => "R10_DATA".R10.AO)
   END_RUNG
   RUNG wire#powerrail
      Contact( "R10_DATA".R10.COOL_RUNNING )
      S_Coil( "R10_RMAP_CV_CONTROL".Config.InvertControl )
   END_RUNG
   RUNG wire#powerrail
      I_Contact( "R10_DATA".R10.COOL_RUNNING )
      R_Coil( "R10_RMAP_CV_CONTROL".Config.InvertControl )
   END_RUNG
   // the same network as SCL:
   #_w1 := "AlwaysTRUE";
   IF "AlwaysTRUE" AND "R10_DATA".R10.RUNNING AND "Valves Data"."A/M".R10 THEN
       "R10_RMAP_CV_CONTROL"(Setpoint := "AO_OUTPUTS"."A/GLR_010_TCV_651_CVOUT",   // PID_Compact
                             Input := "R10_DATA".R10.R10_ramp_substitute,
                             Output_PER => "R10_DATA".R10.AO);
   END_IF;
   "R10_RMAP_CV_CONTROL".Reset := #_w1 AND NOT "R10_DATA".R10.RUNNING;
   IF "R10_RMAP_CV_CONTROL".Reset AND NOT "AlwaysTRUE" THEN
       "A/GLR_010_TCV_651_CVOUT" := 0;
       "R10_DATA".R10.AO := 0;
   END_IF;
   IF "R10_DATA".R10.COOL_RUNNING THEN "R10_RMAP_CV_CONTROL".Config.InvertControl := TRUE; END_IF;
   IF NOT "R10_DATA".R10.COOL_RUNNING THEN "R10_RMAP_CV_CONTROL".Config.InvertControl := FALSE; END_IF;
END_REGION

REGION Network 71: R10 SCADA OUTPUT
   RUNG wire#powerrail
      Contact( "AlwaysTRUE" )
      { S7_Templates := "[SrcType := Int, DestType := Real]" } Normalize(min := "R10_DATA".R10.NORM_MIN, value := "R10_DATA".R10.AO, max := "R10_DATA".R10.NORM_MAX, out => "R10_DATA".R10.NORM_OUT)
      { S7_Templates := "[SrcType := Real, DestType := Real]" } Scale(min := "R10_DATA".R10.SCALE_MIN, value := "R10_DATA".R10.NORM_OUT, max := "R10_DATA".R10.SCALE_MAX, out => "R10_DATA".R10.SCVOUT)
   END_RUNG
   // the same network as SCL:
   IF "AlwaysTRUE" THEN
       "R10_DATA".R10.NORM_OUT := NORM_X(MIN := "R10_DATA".R10.NORM_MIN, VALUE := "R10_DATA".R10.AO, MAX := "R10_DATA".R10.NORM_MAX);
       "R10_DATA".R10.SCVOUT := SCALE_X(MIN := "R10_DATA".R10.SCALE_MIN, VALUE := "R10_DATA".R10.NORM_OUT, MAX := "R10_DATA".R10.SCALE_MAX);
   END_IF;
END_REGION

REGION Network 72: R10 AUTO/MANUAL OUTPUT
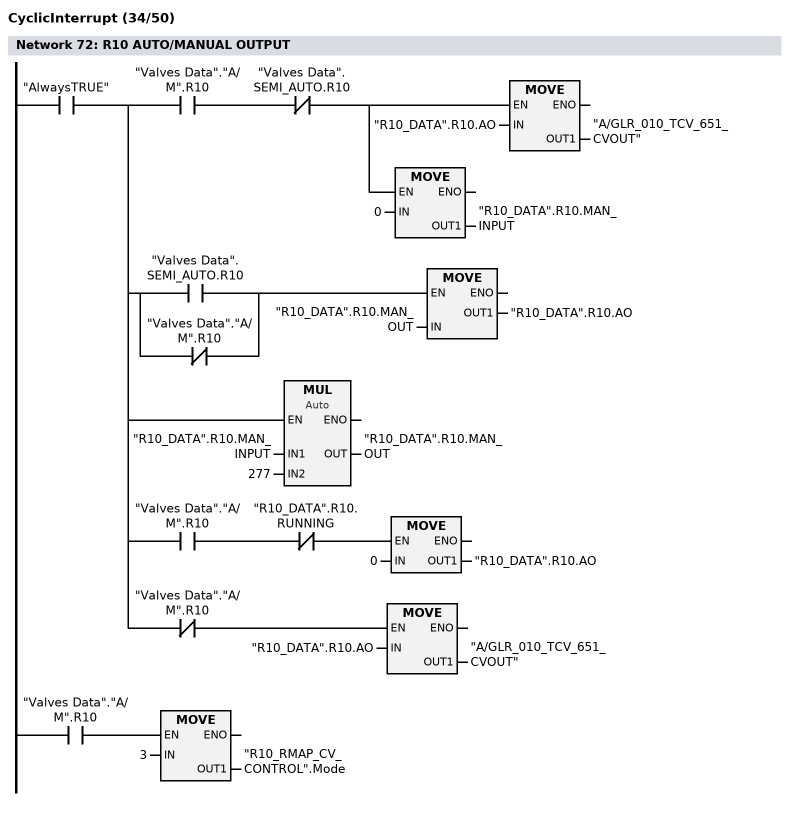
   RUNG wire#powerrail
      Contact( "AlwaysTRUE" )
      wire#w1
      Contact( "Valves Data"."A/M".R10 )
      I_Contact( "Valves Data".SEMI_AUTO.R10 )
      wire#w2
      Move(in := "R10_DATA".R10.AO, out1 => "A/GLR_010_TCV_651_CVOUT")
   END_RUNG
   RUNG wire#w2
      Move(in := 0, out1 => "R10_DATA".R10.MAN_INPUT)
   END_RUNG
   RUNG wire#w1
      Contact( "Valves Data".SEMI_AUTO.R10 )
      wire#w3
      Move(in := "R10_DATA".R10.MAN_OUT, out1 => "R10_DATA".R10.AO)
   END_RUNG
   RUNG wire#w1
      I_Contact( "Valves Data"."A/M".R10 )
   END_RUNG wire#w3
   RUNG wire#w1
      Mul(in1 := "R10_DATA".R10.MAN_INPUT, in2 := 277, out => "R10_DATA".R10.MAN_OUT)
   END_RUNG
   RUNG wire#w1
      Contact( "Valves Data"."A/M".R10 )
      I_Contact( "R10_DATA".R10.RUNNING )
      Move(in := 0, out1 => "R10_DATA".R10.AO)
   END_RUNG
   RUNG wire#w1
      I_Contact( "Valves Data"."A/M".R10 )
      Move(in := "R10_DATA".R10.AO, out1 => "A/GLR_010_TCV_651_CVOUT")
   END_RUNG
   RUNG wire#powerrail
      Contact( "Valves Data"."A/M".R10 )
      Move(in := 3, out1 => "R10_RMAP_CV_CONTROL".Mode)
   END_RUNG
   // the same network as SCL:
   IF "AlwaysTRUE" AND "Valves Data"."A/M".R10 AND NOT "Valves Data".SEMI_AUTO.R10 THEN
       "A/GLR_010_TCV_651_CVOUT" := "R10_DATA".R10.AO;
       "R10_DATA".R10.MAN_INPUT := 0;
   END_IF;
   IF "AlwaysTRUE" AND ("Valves Data".SEMI_AUTO.R10 OR NOT "Valves Data"."A/M".R10) THEN
       "R10_DATA".R10.AO := "R10_DATA".R10.MAN_OUT;
   END_IF;
   IF "AlwaysTRUE" THEN "R10_DATA".R10.MAN_OUT := "R10_DATA".R10.MAN_INPUT * 277; END_IF;
   IF "AlwaysTRUE" AND "Valves Data"."A/M".R10 AND NOT "R10_DATA".R10.RUNNING THEN
       "R10_DATA".R10.AO := 0;
   END_IF;
   IF "AlwaysTRUE" AND NOT "Valves Data"."A/M".R10 THEN
       "A/GLR_010_TCV_651_CVOUT" := "R10_DATA".R10.AO;
   END_IF;
   IF "Valves Data"."A/M".R10 THEN "R10_RMAP_CV_CONTROL".Mode := 3; END_IF;
END_REGION

REGION Network 73: R11_RAMP_CV
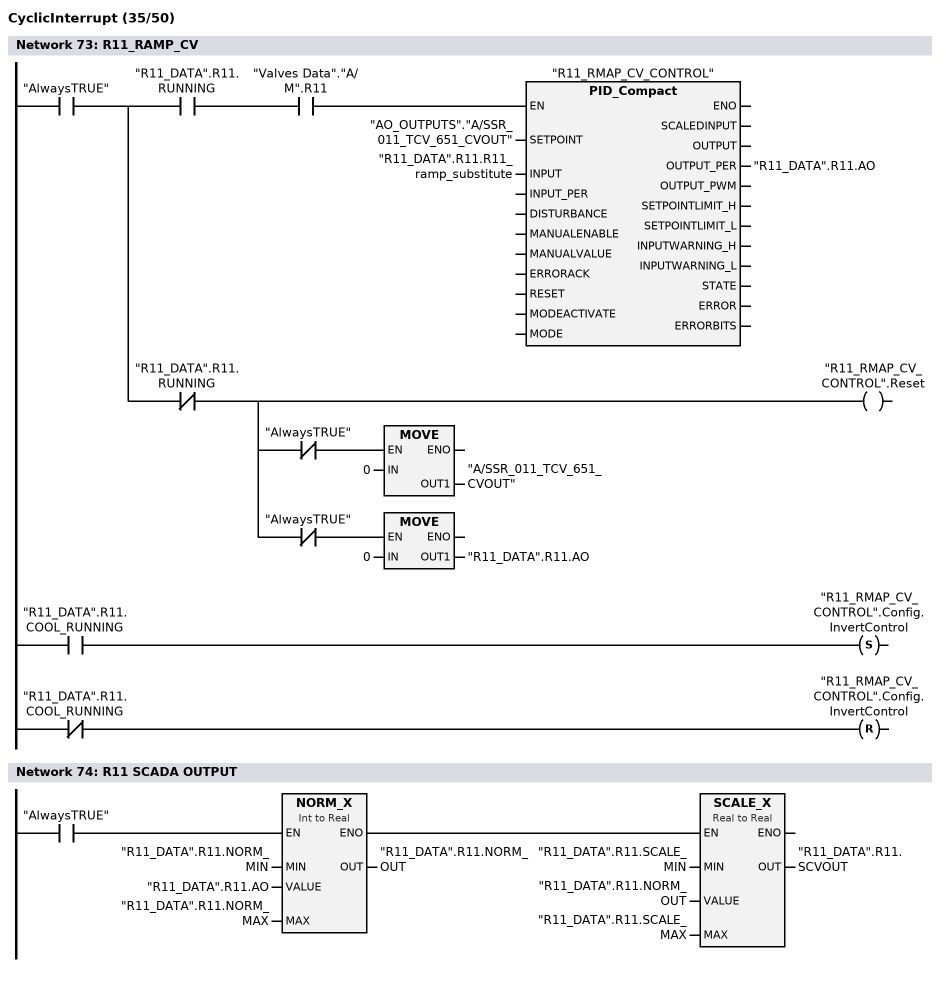
   RUNG wire#powerrail
      Contact( "AlwaysTRUE" )
      wire#w1
      Contact( "R11_DATA".R11.RUNNING )
      Contact( "Valves Data"."A/M".R11 )
      "R11_RMAP_CV_CONTROL".PID_Compact(Setpoint := "AO_OUTPUTS"."A/SSR_011_TCV_651_CVOUT", Input := "R11_DATA".R11.R11_ramp_substitute, Input_PER :=, Disturbance :=, ManualEnable :=, ManualValue :=, ErrorAck :=, Reset :=, ModeActivate :=, Mode :=, ScaledInput =>, Output =>, Output_PER => "R11_DATA".R11.AO, Output_PWM =>, SetpointLimit_H =>, SetpointLimit_L =>, InputWarning_H =>, InputWarning_L =>, State =>, Error =>, ErrorBits =>)
   END_RUNG
   RUNG wire#w1
      I_Contact( "R11_DATA".R11.RUNNING )
      wire#w2
      Coil( "R11_RMAP_CV_CONTROL".Reset )
   END_RUNG
   RUNG wire#w2
      I_Contact( "AlwaysTRUE" )
      Move(in := 0, out1 => "A/SSR_011_TCV_651_CVOUT")
   END_RUNG
   RUNG wire#w2
      I_Contact( "AlwaysTRUE" )
      Move(in := 0, out1 => "R11_DATA".R11.AO)
   END_RUNG
   RUNG wire#powerrail
      Contact( "R11_DATA".R11.COOL_RUNNING )
      S_Coil( "R11_RMAP_CV_CONTROL".Config.InvertControl )
   END_RUNG
   RUNG wire#powerrail
      I_Contact( "R11_DATA".R11.COOL_RUNNING )
      R_Coil( "R11_RMAP_CV_CONTROL".Config.InvertControl )
   END_RUNG
   // the same network as SCL:
   #_w1 := "AlwaysTRUE";
   IF "AlwaysTRUE" AND "R11_DATA".R11.RUNNING AND "Valves Data"."A/M".R11 THEN
       "R11_RMAP_CV_CONTROL"(Setpoint := "AO_OUTPUTS"."A/SSR_011_TCV_651_CVOUT",   // PID_Compact
                             Input := "R11_DATA".R11.R11_ramp_substitute,
                             Output_PER => "R11_DATA".R11.AO);
   END_IF;
   "R11_RMAP_CV_CONTROL".Reset := #_w1 AND NOT "R11_DATA".R11.RUNNING;
   IF "R11_RMAP_CV_CONTROL".Reset AND NOT "AlwaysTRUE" THEN
       "A/SSR_011_TCV_651_CVOUT" := 0;
       "R11_DATA".R11.AO := 0;
   END_IF;
   IF "R11_DATA".R11.COOL_RUNNING THEN "R11_RMAP_CV_CONTROL".Config.InvertControl := TRUE; END_IF;
   IF NOT "R11_DATA".R11.COOL_RUNNING THEN "R11_RMAP_CV_CONTROL".Config.InvertControl := FALSE; END_IF;
END_REGION

REGION Network 74: R11 SCADA OUTPUT
   RUNG wire#powerrail
      Contact( "AlwaysTRUE" )
      { S7_Templates := "[SrcType := Int, DestType := Real]" } Normalize(min := "R11_DATA".R11.NORM_MIN, value := "R11_DATA".R11.AO, max := "R11_DATA".R11.NORM_MAX, out => "R11_DATA".R11.NORM_OUT)
      { S7_Templates := "[SrcType := Real, DestType := Real]" } Scale(min := "R11_DATA".R11.SCALE_MIN, value := "R11_DATA".R11.NORM_OUT, max := "R11_DATA".R11.SCALE_MAX, out => "R11_DATA".R11.SCVOUT)
   END_RUNG
   // the same network as SCL:
   IF "AlwaysTRUE" THEN
       "R11_DATA".R11.NORM_OUT := NORM_X(MIN := "R11_DATA".R11.NORM_MIN, VALUE := "R11_DATA".R11.AO, MAX := "R11_DATA".R11.NORM_MAX);
       "R11_DATA".R11.SCVOUT := SCALE_X(MIN := "R11_DATA".R11.SCALE_MIN, VALUE := "R11_DATA".R11.NORM_OUT, MAX := "R11_DATA".R11.SCALE_MAX);
   END_IF;
END_REGION

REGION Network 75: R11 AUTO/MANUAL OUTPUT
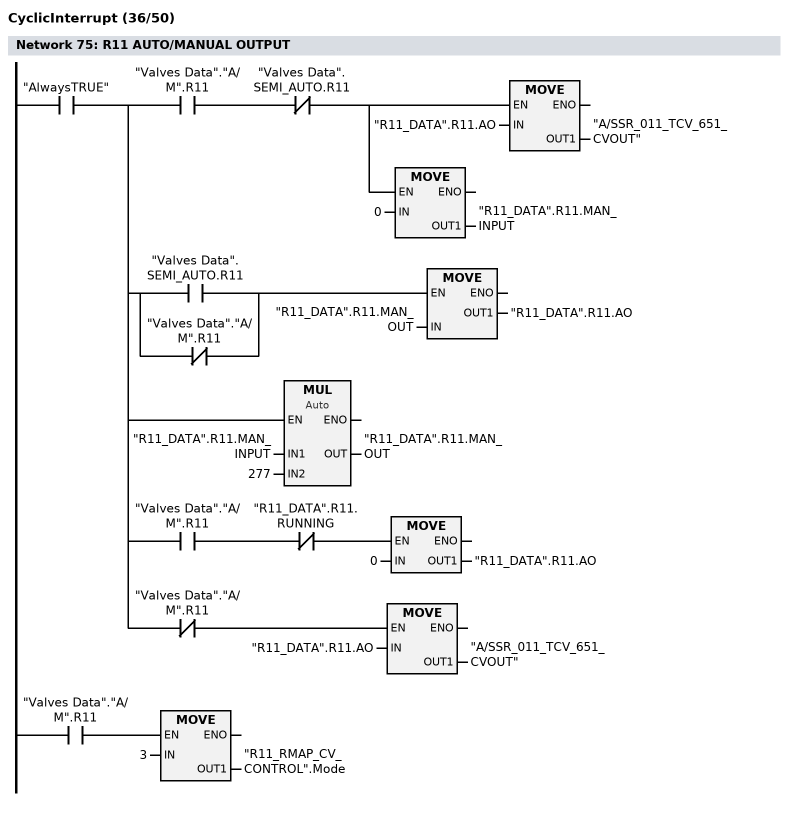
   RUNG wire#powerrail
      Contact( "AlwaysTRUE" )
      wire#w1
      Contact( "Valves Data"."A/M".R11 )
      I_Contact( "Valves Data".SEMI_AUTO.R11 )
      wire#w2
      Move(in := "R11_DATA".R11.AO, out1 => "A/SSR_011_TCV_651_CVOUT")
   END_RUNG
   RUNG wire#w2
      Move(in := 0, out1 => "R11_DATA".R11.MAN_INPUT)
   END_RUNG
   RUNG wire#w1
      Contact( "Valves Data".SEMI_AUTO.R11 )
      wire#w3
      Move(in := "R11_DATA".R11.MAN_OUT, out1 => "R11_DATA".R11.AO)
   END_RUNG
   RUNG wire#w1
      I_Contact( "Valves Data"."A/M".R11 )
   END_RUNG wire#w3
   RUNG wire#w1
      Mul(in1 := "R11_DATA".R11.MAN_INPUT, in2 := 277, out => "R11_DATA".R11.MAN_OUT)
   END_RUNG
   RUNG wire#w1
      Contact( "Valves Data"."A/M".R11 )
      I_Contact( "R11_DATA".R11.RUNNING )
      Move(in := 0, out1 => "R11_DATA".R11.AO)
   END_RUNG
   RUNG wire#w1
      I_Contact( "Valves Data"."A/M".R11 )
      Move(in := "R11_DATA".R11.AO, out1 => "A/SSR_011_TCV_651_CVOUT")
   END_RUNG
   RUNG wire#powerrail
      Contact( "Valves Data"."A/M".R11 )
      Move(in := 3, out1 => "R11_RMAP_CV_CONTROL".Mode)
   END_RUNG
   // the same network as SCL:
   IF "AlwaysTRUE" AND "Valves Data"."A/M".R11 AND NOT "Valves Data".SEMI_AUTO.R11 THEN
       "A/SSR_011_TCV_651_CVOUT" := "R11_DATA".R11.AO;
       "R11_DATA".R11.MAN_INPUT := 0;
   END_IF;
   IF "AlwaysTRUE" AND ("Valves Data".SEMI_AUTO.R11 OR NOT "Valves Data"."A/M".R11) THEN
       "R11_DATA".R11.AO := "R11_DATA".R11.MAN_OUT;
   END_IF;
   IF "AlwaysTRUE" THEN "R11_DATA".R11.MAN_OUT := "R11_DATA".R11.MAN_INPUT * 277; END_IF;
   IF "AlwaysTRUE" AND "Valves Data"."A/M".R11 AND NOT "R11_DATA".R11.RUNNING THEN
       "R11_DATA".R11.AO := 0;
   END_IF;
   IF "AlwaysTRUE" AND NOT "Valves Data"."A/M".R11 THEN
       "A/SSR_011_TCV_651_CVOUT" := "R11_DATA".R11.AO;
   END_IF;
   IF "Valves Data"."A/M".R11 THEN "R11_RMAP_CV_CONTROL".Mode := 3; END_IF;
END_REGION

REGION Network 76: R12_RAMP_CV
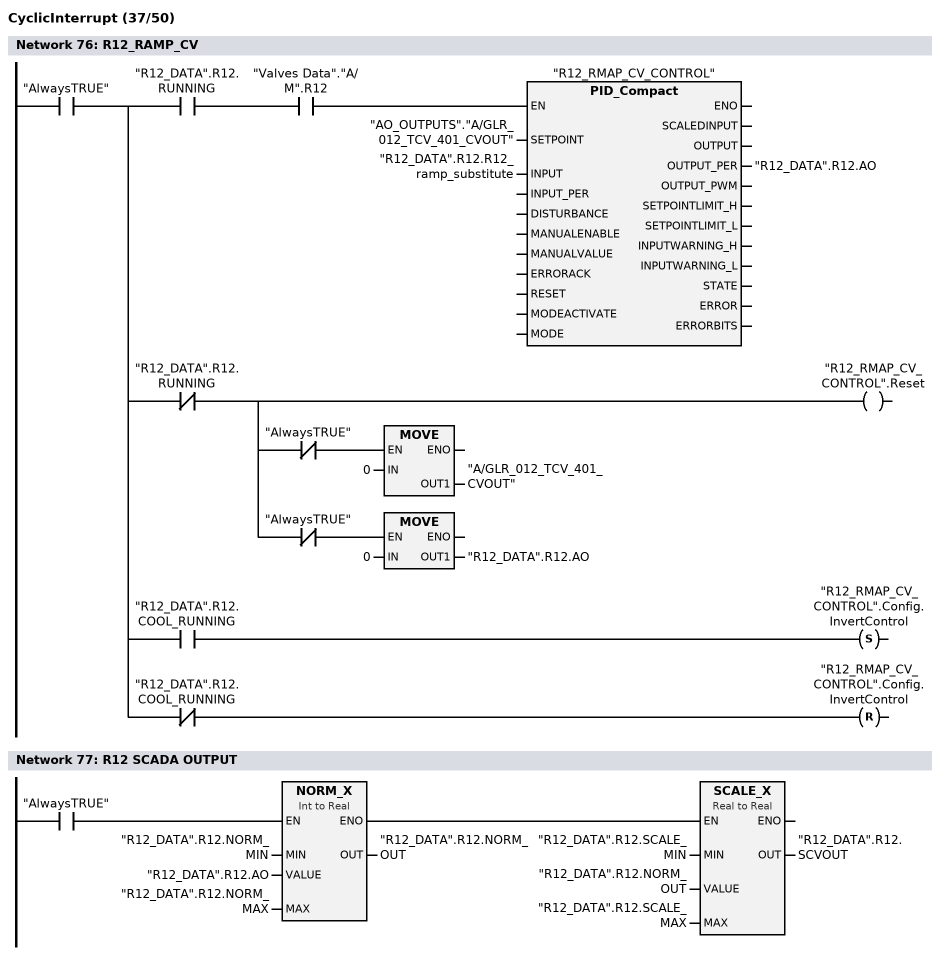
   RUNG wire#powerrail
      Contact( "AlwaysTRUE" )
      wire#w1
      Contact( "R12_DATA".R12.RUNNING )
      Contact( "Valves Data"."A/M".R12 )
      "R12_RMAP_CV_CONTROL".PID_Compact(Setpoint := "AO_OUTPUTS"."A/GLR_012_TCV_401_CVOUT", Input := "R12_DATA".R12.R12_ramp_substitute, Input_PER :=, Disturbance :=, ManualEnable :=, ManualValue :=, ErrorAck :=, Reset :=, ModeActivate :=, Mode :=, ScaledInput =>, Output =>, Output_PER => "R12_DATA".R12.AO, Output_PWM =>, SetpointLimit_H =>, SetpointLimit_L =>, InputWarning_H =>, InputWarning_L =>, State =>, Error =>, ErrorBits =>)
   END_RUNG
   RUNG wire#w1
      I_Contact( "R12_DATA".R12.RUNNING )
      wire#w2
      Coil( "R12_RMAP_CV_CONTROL".Reset )
   END_RUNG
   RUNG wire#w2
      I_Contact( "AlwaysTRUE" )
      Move(in := 0, out1 => "A/GLR_012_TCV_401_CVOUT")
   END_RUNG
   RUNG wire#w2
      I_Contact( "AlwaysTRUE" )
      Move(in := 0, out1 => "R12_DATA".R12.AO)
   END_RUNG
   RUNG wire#w1
      Contact( "R12_DATA".R12.COOL_RUNNING )
      S_Coil( "R12_RMAP_CV_CONTROL".Config.InvertControl )
   END_RUNG
   RUNG wire#w1
      I_Contact( "R12_DATA".R12.COOL_RUNNING )
      R_Coil( "R12_RMAP_CV_CONTROL".Config.InvertControl )
   END_RUNG
   // the same network as SCL:
   #_w1 := "AlwaysTRUE";
   IF "AlwaysTRUE" AND "R12_DATA".R12.RUNNING AND "Valves Data"."A/M".R12 THEN
       "R12_RMAP_CV_CONTROL"(Setpoint := "AO_OUTPUTS"."A/GLR_012_TCV_401_CVOUT",   // PID_Compact
                             Input := "R12_DATA".R12.R12_ramp_substitute,
                             Output_PER => "R12_DATA".R12.AO);
   END_IF;
   "R12_RMAP_CV_CONTROL".Reset := #_w1 AND NOT "R12_DATA".R12.RUNNING;
   IF "R12_RMAP_CV_CONTROL".Reset AND NOT "AlwaysTRUE" THEN
       "A/GLR_012_TCV_401_CVOUT" := 0;
       "R12_DATA".R12.AO := 0;
   END_IF;
   IF #_w1 AND "R12_DATA".R12.COOL_RUNNING THEN "R12_RMAP_CV_CONTROL".Config.InvertControl := TRUE; END_IF;
   IF #_w1 AND NOT "R12_DATA".R12.COOL_RUNNING THEN
       "R12_RMAP_CV_CONTROL".Config.InvertControl := FALSE;
   END_IF;
END_REGION

REGION Network 77: R12 SCADA OUTPUT
   RUNG wire#powerrail
      Contact( "AlwaysTRUE" )
      { S7_Templates := "[SrcType := Int, DestType := Real]" } Normalize(min := "R12_DATA".R12.NORM_MIN, value := "R12_DATA".R12.AO, max := "R12_DATA".R12.NORM_MAX, out => "R12_DATA".R12.NORM_OUT)
      { S7_Templates := "[SrcType := Real, DestType := Real]" } Scale(min := "R12_DATA".R12.SCALE_MIN, value := "R12_DATA".R12.NORM_OUT, max := "R12_DATA".R12.SCALE_MAX, out => "R12_DATA".R12.SCVOUT)
   END_RUNG
   // the same network as SCL:
   IF "AlwaysTRUE" THEN
       "R12_DATA".R12.NORM_OUT := NORM_X(MIN := "R12_DATA".R12.NORM_MIN, VALUE := "R12_DATA".R12.AO, MAX := "R12_DATA".R12.NORM_MAX);
       "R12_DATA".R12.SCVOUT := SCALE_X(MIN := "R12_DATA".R12.SCALE_MIN, VALUE := "R12_DATA".R12.NORM_OUT, MAX := "R12_DATA".R12.SCALE_MAX);
   END_IF;
END_REGION

REGION Network 78: R12 AUTO/MANUAL OUTPUT
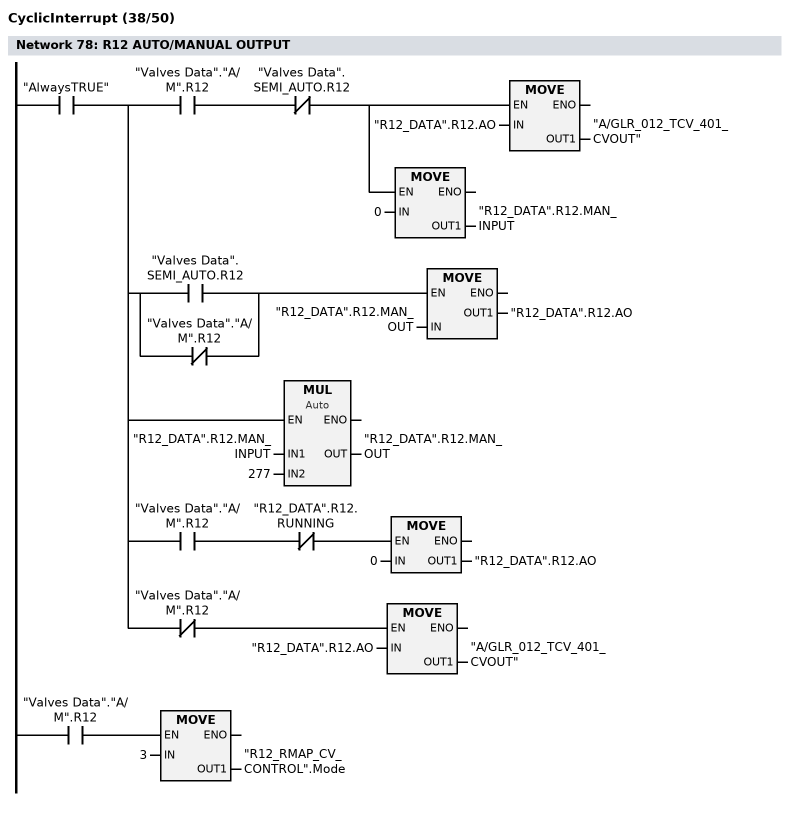
   RUNG wire#powerrail
      Contact( "AlwaysTRUE" )
      wire#w1
      Contact( "Valves Data"."A/M".R12 )
      I_Contact( "Valves Data".SEMI_AUTO.R12 )
      wire#w2
      Move(in := "R12_DATA".R12.AO, out1 => "A/GLR_012_TCV_401_CVOUT")
   END_RUNG
   RUNG wire#w2
      Move(in := 0, out1 => "R12_DATA".R12.MAN_INPUT)
   END_RUNG
   RUNG wire#w1
      Contact( "Valves Data".SEMI_AUTO.R12 )
      wire#w3
      Move(in := "R12_DATA".R12.MAN_OUT, out1 => "R12_DATA".R12.AO)
   END_RUNG
   RUNG wire#w1
      I_Contact( "Valves Data"."A/M".R12 )
   END_RUNG wire#w3
   RUNG wire#w1
      Mul(in1 := "R12_DATA".R12.MAN_INPUT, in2 := 277, out => "R12_DATA".R12.MAN_OUT)
   END_RUNG
   RUNG wire#w1
      Contact( "Valves Data"."A/M".R12 )
      I_Contact( "R12_DATA".R12.RUNNING )
      Move(in := 0, out1 => "R12_DATA".R12.AO)
   END_RUNG
   RUNG wire#w1
      I_Contact( "Valves Data"."A/M".R12 )
      Move(in := "R12_DATA".R12.AO, out1 => "A/GLR_012_TCV_401_CVOUT")
   END_RUNG
   RUNG wire#powerrail
      Contact( "Valves Data"."A/M".R12 )
      Move(in := 3, out1 => "R12_RMAP_CV_CONTROL".Mode)
   END_RUNG
   // the same network as SCL:
   IF "AlwaysTRUE" AND "Valves Data"."A/M".R12 AND NOT "Valves Data".SEMI_AUTO.R12 THEN
       "A/GLR_012_TCV_401_CVOUT" := "R12_DATA".R12.AO;
       "R12_DATA".R12.MAN_INPUT := 0;
   END_IF;
   IF "AlwaysTRUE" AND ("Valves Data".SEMI_AUTO.R12 OR NOT "Valves Data"."A/M".R12) THEN
       "R12_DATA".R12.AO := "R12_DATA".R12.MAN_OUT;
   END_IF;
   IF "AlwaysTRUE" THEN "R12_DATA".R12.MAN_OUT := "R12_DATA".R12.MAN_INPUT * 277; END_IF;
   IF "AlwaysTRUE" AND "Valves Data"."A/M".R12 AND NOT "R12_DATA".R12.RUNNING THEN
       "R12_DATA".R12.AO := 0;
   END_IF;
   IF "AlwaysTRUE" AND NOT "Valves Data"."A/M".R12 THEN
       "A/GLR_012_TCV_401_CVOUT" := "R12_DATA".R12.AO;
   END_IF;
   IF "Valves Data"."A/M".R12 THEN "R12_RMAP_CV_CONTROL".Mode := 3; END_IF;
END_REGION

REGION Network 79: R13_RAMP_CV
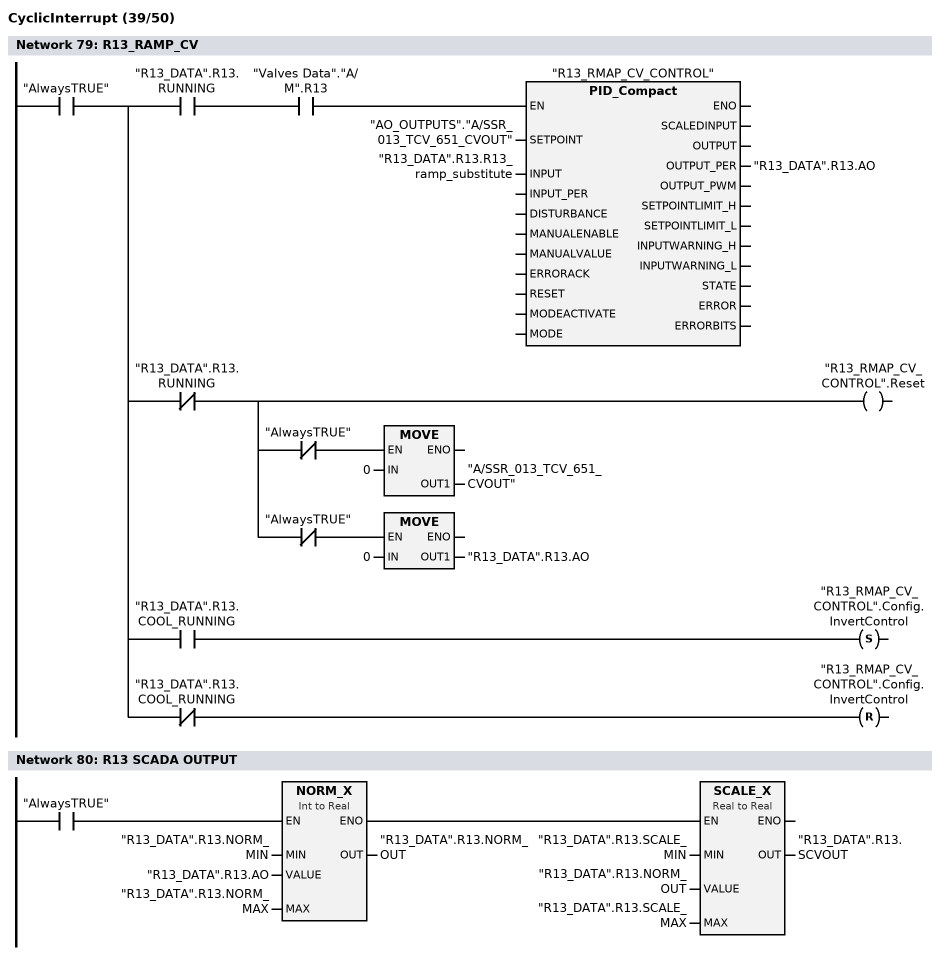
   RUNG wire#powerrail
      Contact( "AlwaysTRUE" )
      wire#w1
      Contact( "R13_DATA".R13.RUNNING )
      Contact( "Valves Data"."A/M".R13 )
      "R13_RMAP_CV_CONTROL".PID_Compact(Setpoint := "AO_OUTPUTS"."A/SSR_013_TCV_651_CVOUT", Input := "R13_DATA".R13.R13_ramp_substitute, Input_PER :=, Disturbance :=, ManualEnable :=, ManualValue :=, ErrorAck :=, Reset :=, ModeActivate :=, Mode :=, ScaledInput =>, Output =>, Output_PER => "R13_DATA".R13.AO, Output_PWM =>, SetpointLimit_H =>, SetpointLimit_L =>, InputWarning_H =>, InputWarning_L =>, State =>, Error =>, ErrorBits =>)
   END_RUNG
   RUNG wire#w1
      I_Contact( "R13_DATA".R13.RUNNING )
      wire#w2
      Coil( "R13_RMAP_CV_CONTROL".Reset )
   END_RUNG
   RUNG wire#w2
      I_Contact( "AlwaysTRUE" )
      Move(in := 0, out1 => "A/SSR_013_TCV_651_CVOUT")
   END_RUNG
   RUNG wire#w2
      I_Contact( "AlwaysTRUE" )
      Move(in := 0, out1 => "R13_DATA".R13.AO)
   END_RUNG
   RUNG wire#w1
      Contact( "R13_DATA".R13.COOL_RUNNING )
      S_Coil( "R13_RMAP_CV_CONTROL".Config.InvertControl )
   END_RUNG
   RUNG wire#w1
      I_Contact( "R13_DATA".R13.COOL_RUNNING )
      R_Coil( "R13_RMAP_CV_CONTROL".Config.InvertControl )
   END_RUNG
   // the same network as SCL:
   #_w1 := "AlwaysTRUE";
   IF "AlwaysTRUE" AND "R13_DATA".R13.RUNNING AND "Valves Data"."A/M".R13 THEN
       "R13_RMAP_CV_CONTROL"(Setpoint := "AO_OUTPUTS"."A/SSR_013_TCV_651_CVOUT",   // PID_Compact
                             Input := "R13_DATA".R13.R13_ramp_substitute,
                             Output_PER => "R13_DATA".R13.AO);
   END_IF;
   "R13_RMAP_CV_CONTROL".Reset := #_w1 AND NOT "R13_DATA".R13.RUNNING;
   IF "R13_RMAP_CV_CONTROL".Reset AND NOT "AlwaysTRUE" THEN
       "A/SSR_013_TCV_651_CVOUT" := 0;
       "R13_DATA".R13.AO := 0;
   END_IF;
   IF #_w1 AND "R13_DATA".R13.COOL_RUNNING THEN "R13_RMAP_CV_CONTROL".Config.InvertControl := TRUE; END_IF;
   IF #_w1 AND NOT "R13_DATA".R13.COOL_RUNNING THEN
       "R13_RMAP_CV_CONTROL".Config.InvertControl := FALSE;
   END_IF;
END_REGION

REGION Network 80: R13 SCADA OUTPUT
   RUNG wire#powerrail
      Contact( "AlwaysTRUE" )
      { S7_Templates := "[SrcType := Int, DestType := Real]" } Normalize(min := "R13_DATA".R13.NORM_MIN, value := "R13_DATA".R13.AO, max := "R13_DATA".R13.NORM_MAX, out => "R13_DATA".R13.NORM_OUT)
      { S7_Templates := "[SrcType := Real, DestType := Real]" } Scale(min := "R13_DATA".R13.SCALE_MIN, value := "R13_DATA".R13.NORM_OUT, max := "R13_DATA".R13.SCALE_MAX, out => "R13_DATA".R13.SCVOUT)
   END_RUNG
   // the same network as SCL:
   IF "AlwaysTRUE" THEN
       "R13_DATA".R13.NORM_OUT := NORM_X(MIN := "R13_DATA".R13.NORM_MIN, VALUE := "R13_DATA".R13.AO, MAX := "R13_DATA".R13.NORM_MAX);
       "R13_DATA".R13.SCVOUT := SCALE_X(MIN := "R13_DATA".R13.SCALE_MIN, VALUE := "R13_DATA".R13.NORM_OUT, MAX := "R13_DATA".R13.SCALE_MAX);
   END_IF;
END_REGION

REGION Network 81: R13 AUTO/MANUAL OUTPUT
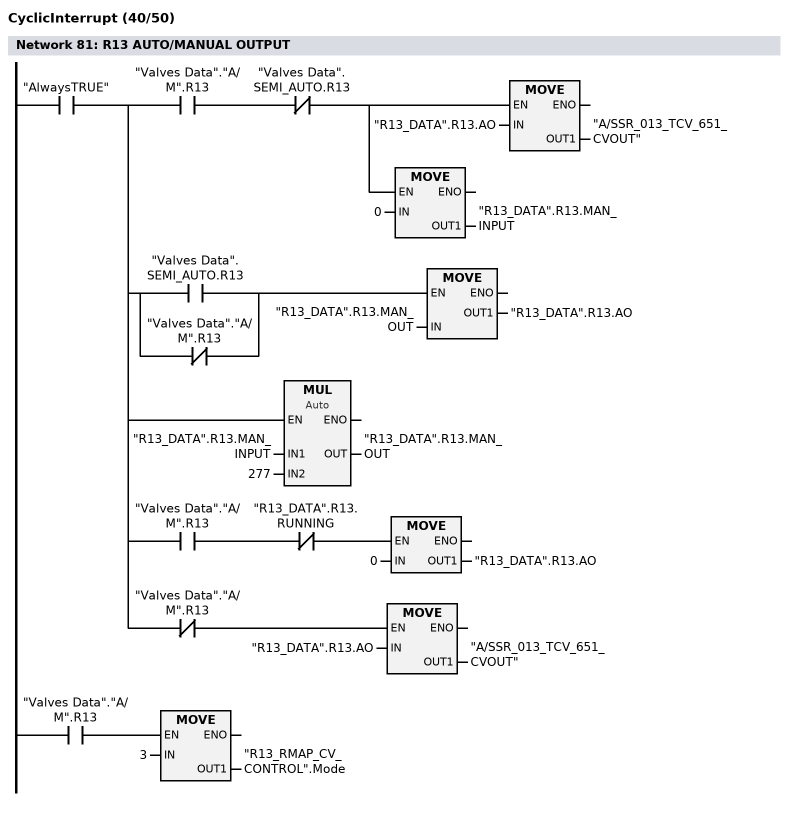
   RUNG wire#powerrail
      Contact( "AlwaysTRUE" )
      wire#w1
      Contact( "Valves Data"."A/M".R13 )
      I_Contact( "Valves Data".SEMI_AUTO.R13 )
      wire#w2
      Move(in := "R13_DATA".R13.AO, out1 => "A/SSR_013_TCV_651_CVOUT")
   END_RUNG
   RUNG wire#w2
      Move(in := 0, out1 => "R13_DATA".R13.MAN_INPUT)
   END_RUNG
   RUNG wire#w1
      Contact( "Valves Data".SEMI_AUTO.R13 )
      wire#w3
      Move(in := "R13_DATA".R13.MAN_OUT, out1 => "R13_DATA".R13.AO)
   END_RUNG
   RUNG wire#w1
      I_Contact( "Valves Data"."A/M".R13 )
   END_RUNG wire#w3
   RUNG wire#w1
      Mul(in1 := "R13_DATA".R13.MAN_INPUT, in2 := 277, out => "R13_DATA".R13.MAN_OUT)
   END_RUNG
   RUNG wire#w1
      Contact( "Valves Data"."A/M".R13 )
      I_Contact( "R13_DATA".R13.RUNNING )
      Move(in := 0, out1 => "R13_DATA".R13.AO)
   END_RUNG
   RUNG wire#w1
      I_Contact( "Valves Data"."A/M".R13 )
      Move(in := "R13_DATA".R13.AO, out1 => "A/SSR_013_TCV_651_CVOUT")
   END_RUNG
   RUNG wire#powerrail
      Contact( "Valves Data"."A/M".R13 )
      Move(in := 3, out1 => "R13_RMAP_CV_CONTROL".Mode)
   END_RUNG
   // the same network as SCL:
   IF "AlwaysTRUE" AND "Valves Data"."A/M".R13 AND NOT "Valves Data".SEMI_AUTO.R13 THEN
       "A/SSR_013_TCV_651_CVOUT" := "R13_DATA".R13.AO;
       "R13_DATA".R13.MAN_INPUT := 0;
   END_IF;
   IF "AlwaysTRUE" AND ("Valves Data".SEMI_AUTO.R13 OR NOT "Valves Data"."A/M".R13) THEN
       "R13_DATA".R13.AO := "R13_DATA".R13.MAN_OUT;
   END_IF;
   IF "AlwaysTRUE" THEN "R13_DATA".R13.MAN_OUT := "R13_DATA".R13.MAN_INPUT * 277; END_IF;
   IF "AlwaysTRUE" AND "Valves Data"."A/M".R13 AND NOT "R13_DATA".R13.RUNNING THEN
       "R13_DATA".R13.AO := 0;
   END_IF;
   IF "AlwaysTRUE" AND NOT "Valves Data"."A/M".R13 THEN
       "A/SSR_013_TCV_651_CVOUT" := "R13_DATA".R13.AO;
   END_IF;
   IF "Valves Data"."A/M".R13 THEN "R13_RMAP_CV_CONTROL".Mode := 3; END_IF;
END_REGION

REGION Network 82: R14_RAMP_CV
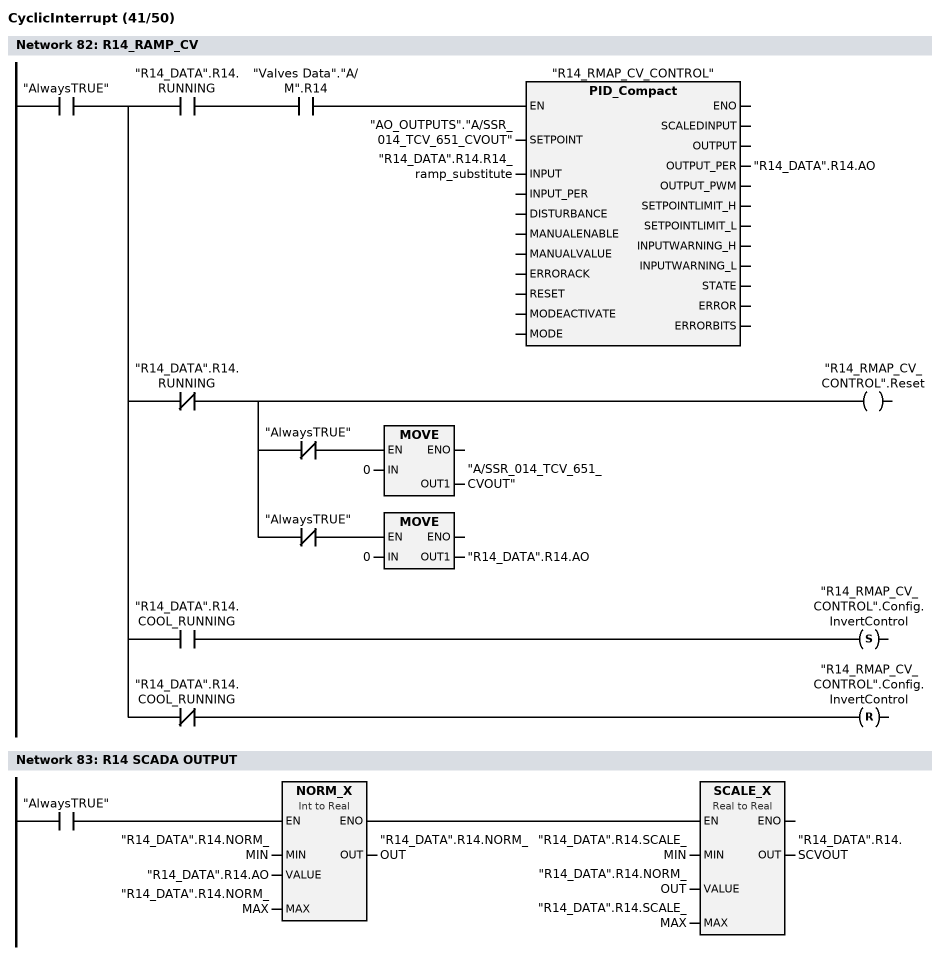
   RUNG wire#powerrail
      Contact( "AlwaysTRUE" )
      wire#w1
      Contact( "R14_DATA".R14.RUNNING )
      Contact( "Valves Data"."A/M".R14 )
      "R14_RMAP_CV_CONTROL".PID_Compact(Setpoint := "AO_OUTPUTS"."A/SSR_014_TCV_651_CVOUT", Input := "R14_DATA".R14.R14_ramp_substitute, Input_PER :=, Disturbance :=, ManualEnable :=, ManualValue :=, ErrorAck :=, Reset :=, ModeActivate :=, Mode :=, ScaledInput =>, Output =>, Output_PER => "R14_DATA".R14.AO, Output_PWM =>, SetpointLimit_H =>, SetpointLimit_L =>, InputWarning_H =>, InputWarning_L =>, State =>, Error =>, ErrorBits =>)
   END_RUNG
   RUNG wire#w1
      I_Contact( "R14_DATA".R14.RUNNING )
      wire#w2
      Coil( "R14_RMAP_CV_CONTROL".Reset )
   END_RUNG
   RUNG wire#w2
      I_Contact( "AlwaysTRUE" )
      Move(in := 0, out1 => "A/SSR_014_TCV_651_CVOUT")
   END_RUNG
   RUNG wire#w2
      I_Contact( "AlwaysTRUE" )
      Move(in := 0, out1 => "R14_DATA".R14.AO)
   END_RUNG
   RUNG wire#w1
      Contact( "R14_DATA".R14.COOL_RUNNING )
      S_Coil( "R14_RMAP_CV_CONTROL".Config.InvertControl )
   END_RUNG
   RUNG wire#w1
      I_Contact( "R14_DATA".R14.COOL_RUNNING )
      R_Coil( "R14_RMAP_CV_CONTROL".Config.InvertControl )
   END_RUNG
   // the same network as SCL:
   #_w1 := "AlwaysTRUE";
   IF "AlwaysTRUE" AND "R14_DATA".R14.RUNNING AND "Valves Data"."A/M".R14 THEN
       "R14_RMAP_CV_CONTROL"(Setpoint := "AO_OUTPUTS"."A/SSR_014_TCV_651_CVOUT",   // PID_Compact
                             Input := "R14_DATA".R14.R14_ramp_substitute,
                             Output_PER => "R14_DATA".R14.AO);
   END_IF;
   "R14_RMAP_CV_CONTROL".Reset := #_w1 AND NOT "R14_DATA".R14.RUNNING;
   IF "R14_RMAP_CV_CONTROL".Reset AND NOT "AlwaysTRUE" THEN
       "A/SSR_014_TCV_651_CVOUT" := 0;
       "R14_DATA".R14.AO := 0;
   END_IF;
   IF #_w1 AND "R14_DATA".R14.COOL_RUNNING THEN "R14_RMAP_CV_CONTROL".Config.InvertControl := TRUE; END_IF;
   IF #_w1 AND NOT "R14_DATA".R14.COOL_RUNNING THEN
       "R14_RMAP_CV_CONTROL".Config.InvertControl := FALSE;
   END_IF;
END_REGION

REGION Network 83: R14 SCADA OUTPUT
   RUNG wire#powerrail
      Contact( "AlwaysTRUE" )
      { S7_Templates := "[SrcType := Int, DestType := Real]" } Normalize(min := "R14_DATA".R14.NORM_MIN, value := "R14_DATA".R14.AO, max := "R14_DATA".R14.NORM_MAX, out => "R14_DATA".R14.NORM_OUT)
      { S7_Templates := "[SrcType := Real, DestType := Real]" } Scale(min := "R14_DATA".R14.SCALE_MIN, value := "R14_DATA".R14.NORM_OUT, max := "R14_DATA".R14.SCALE_MAX, out => "R14_DATA".R14.SCVOUT)
   END_RUNG
   // the same network as SCL:
   IF "AlwaysTRUE" THEN
       "R14_DATA".R14.NORM_OUT := NORM_X(MIN := "R14_DATA".R14.NORM_MIN, VALUE := "R14_DATA".R14.AO, MAX := "R14_DATA".R14.NORM_MAX);
       "R14_DATA".R14.SCVOUT := SCALE_X(MIN := "R14_DATA".R14.SCALE_MIN, VALUE := "R14_DATA".R14.NORM_OUT, MAX := "R14_DATA".R14.SCALE_MAX);
   END_IF;
END_REGION

REGION Network 84: R14 AUTO/MANUAL OUTPUT
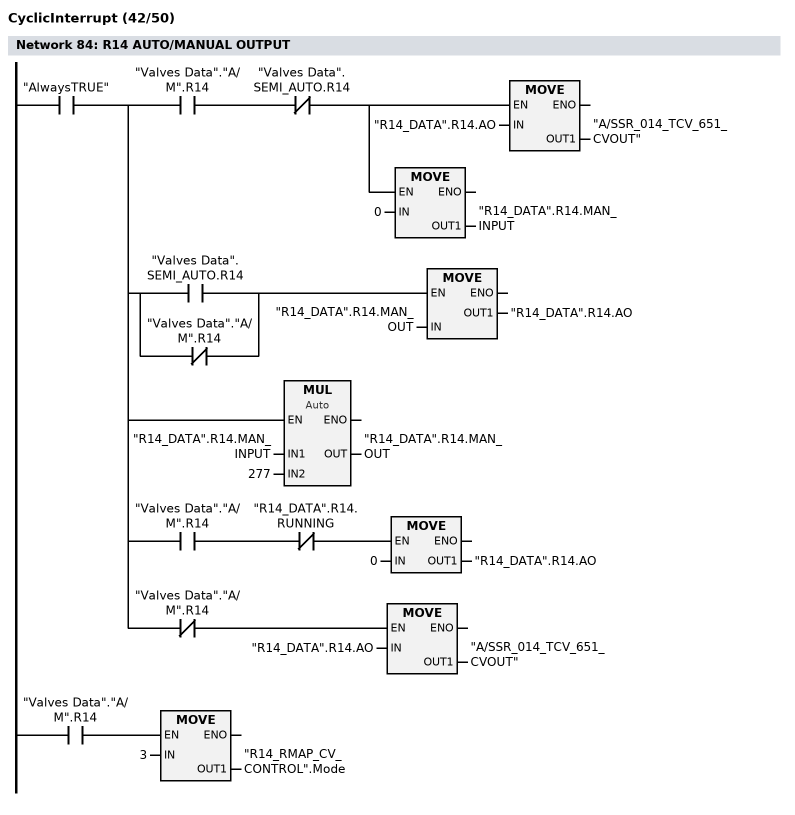
   RUNG wire#powerrail
      Contact( "AlwaysTRUE" )
      wire#w1
      Contact( "Valves Data"."A/M".R14 )
      I_Contact( "Valves Data".SEMI_AUTO.R14 )
      wire#w2
      Move(in := "R14_DATA".R14.AO, out1 => "A/SSR_014_TCV_651_CVOUT")
   END_RUNG
   RUNG wire#w2
      Move(in := 0, out1 => "R14_DATA".R14.MAN_INPUT)
   END_RUNG
   RUNG wire#w1
      Contact( "Valves Data".SEMI_AUTO.R14 )
      wire#w3
      Move(in := "R14_DATA".R14.MAN_OUT, out1 => "R14_DATA".R14.AO)
   END_RUNG
   RUNG wire#w1
      I_Contact( "Valves Data"."A/M".R14 )
   END_RUNG wire#w3
   RUNG wire#w1
      Mul(in1 := "R14_DATA".R14.MAN_INPUT, in2 := 277, out => "R14_DATA".R14.MAN_OUT)
   END_RUNG
   RUNG wire#w1
      Contact( "Valves Data"."A/M".R14 )
      I_Contact( "R14_DATA".R14.RUNNING )
      Move(in := 0, out1 => "R14_DATA".R14.AO)
   END_RUNG
   RUNG wire#w1
      I_Contact( "Valves Data"."A/M".R14 )
      Move(in := "R14_DATA".R14.AO, out1 => "A/SSR_014_TCV_651_CVOUT")
   END_RUNG
   RUNG wire#powerrail
      Contact( "Valves Data"."A/M".R14 )
      Move(in := 3, out1 => "R14_RMAP_CV_CONTROL".Mode)
   END_RUNG
   // the same network as SCL:
   IF "AlwaysTRUE" AND "Valves Data"."A/M".R14 AND NOT "Valves Data".SEMI_AUTO.R14 THEN
       "A/SSR_014_TCV_651_CVOUT" := "R14_DATA".R14.AO;
       "R14_DATA".R14.MAN_INPUT := 0;
   END_IF;
   IF "AlwaysTRUE" AND ("Valves Data".SEMI_AUTO.R14 OR NOT "Valves Data"."A/M".R14) THEN
       "R14_DATA".R14.AO := "R14_DATA".R14.MAN_OUT;
   END_IF;
   IF "AlwaysTRUE" THEN "R14_DATA".R14.MAN_OUT := "R14_DATA".R14.MAN_INPUT * 277; END_IF;
   IF "AlwaysTRUE" AND "Valves Data"."A/M".R14 AND NOT "R14_DATA".R14.RUNNING THEN
       "R14_DATA".R14.AO := 0;
   END_IF;
   IF "AlwaysTRUE" AND NOT "Valves Data"."A/M".R14 THEN
       "A/SSR_014_TCV_651_CVOUT" := "R14_DATA".R14.AO;
   END_IF;
   IF "Valves Data"."A/M".R14 THEN "R14_RMAP_CV_CONTROL".Mode := 3; END_IF;
END_REGION

REGION Network 85: R15_RAMP_CV
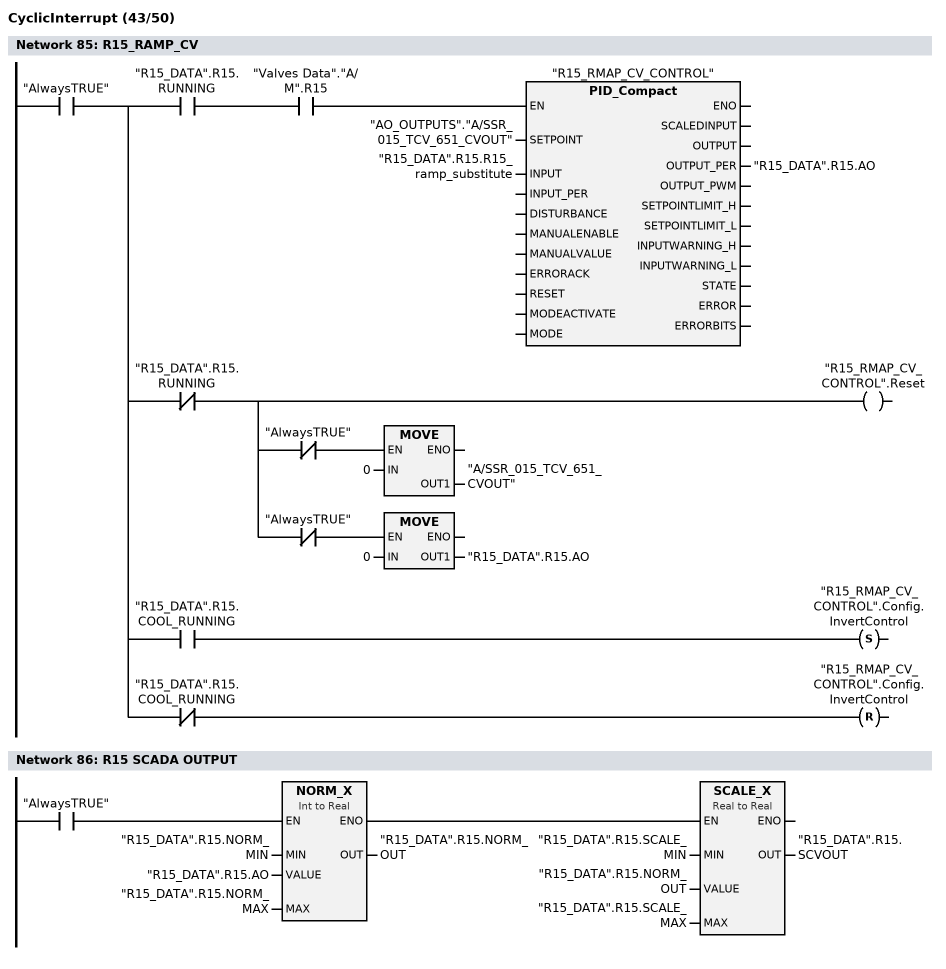
   RUNG wire#powerrail
      Contact( "AlwaysTRUE" )
      wire#w1
      Contact( "R15_DATA".R15.RUNNING )
      Contact( "Valves Data"."A/M".R15 )
      "R15_RMAP_CV_CONTROL".PID_Compact(Setpoint := "AO_OUTPUTS"."A/SSR_015_TCV_651_CVOUT", Input := "R15_DATA".R15.R15_ramp_substitute, Input_PER :=, Disturbance :=, ManualEnable :=, ManualValue :=, ErrorAck :=, Reset :=, ModeActivate :=, Mode :=, ScaledInput =>, Output =>, Output_PER => "R15_DATA".R15.AO, Output_PWM =>, SetpointLimit_H =>, SetpointLimit_L =>, InputWarning_H =>, InputWarning_L =>, State =>, Error =>, ErrorBits =>)
   END_RUNG
   RUNG wire#w1
      I_Contact( "R15_DATA".R15.RUNNING )
      wire#w2
      Coil( "R15_RMAP_CV_CONTROL".Reset )
   END_RUNG
   RUNG wire#w2
      I_Contact( "AlwaysTRUE" )
      Move(in := 0, out1 => "A/SSR_015_TCV_651_CVOUT")
   END_RUNG
   RUNG wire#w2
      I_Contact( "AlwaysTRUE" )
      Move(in := 0, out1 => "R15_DATA".R15.AO)
   END_RUNG
   RUNG wire#w1
      Contact( "R15_DATA".R15.COOL_RUNNING )
      S_Coil( "R15_RMAP_CV_CONTROL".Config.InvertControl )
   END_RUNG
   RUNG wire#w1
      I_Contact( "R15_DATA".R15.COOL_RUNNING )
      R_Coil( "R15_RMAP_CV_CONTROL".Config.InvertControl )
   END_RUNG
   // the same network as SCL:
   #_w1 := "AlwaysTRUE";
   IF "AlwaysTRUE" AND "R15_DATA".R15.RUNNING AND "Valves Data"."A/M".R15 THEN
       "R15_RMAP_CV_CONTROL"(Setpoint := "AO_OUTPUTS"."A/SSR_015_TCV_651_CVOUT",   // PID_Compact
                             Input := "R15_DATA".R15.R15_ramp_substitute,
                             Output_PER => "R15_DATA".R15.AO);
   END_IF;
   "R15_RMAP_CV_CONTROL".Reset := #_w1 AND NOT "R15_DATA".R15.RUNNING;
   IF "R15_RMAP_CV_CONTROL".Reset AND NOT "AlwaysTRUE" THEN
       "A/SSR_015_TCV_651_CVOUT" := 0;
       "R15_DATA".R15.AO := 0;
   END_IF;
   IF #_w1 AND "R15_DATA".R15.COOL_RUNNING THEN "R15_RMAP_CV_CONTROL".Config.InvertControl := TRUE; END_IF;
   IF #_w1 AND NOT "R15_DATA".R15.COOL_RUNNING THEN
       "R15_RMAP_CV_CONTROL".Config.InvertControl := FALSE;
   END_IF;
END_REGION

REGION Network 86: R15 SCADA OUTPUT
   RUNG wire#powerrail
      Contact( "AlwaysTRUE" )
      { S7_Templates := "[SrcType := Int, DestType := Real]" } Normalize(min := "R15_DATA".R15.NORM_MIN, value := "R15_DATA".R15.AO, max := "R15_DATA".R15.NORM_MAX, out => "R15_DATA".R15.NORM_OUT)
      { S7_Templates := "[SrcType := Real, DestType := Real]" } Scale(min := "R15_DATA".R15.SCALE_MIN, value := "R15_DATA".R15.NORM_OUT, max := "R15_DATA".R15.SCALE_MAX, out => "R15_DATA".R15.SCVOUT)
   END_RUNG
   // the same network as SCL:
   IF "AlwaysTRUE" THEN
       "R15_DATA".R15.NORM_OUT := NORM_X(MIN := "R15_DATA".R15.NORM_MIN, VALUE := "R15_DATA".R15.AO, MAX := "R15_DATA".R15.NORM_MAX);
       "R15_DATA".R15.SCVOUT := SCALE_X(MIN := "R15_DATA".R15.SCALE_MIN, VALUE := "R15_DATA".R15.NORM_OUT, MAX := "R15_DATA".R15.SCALE_MAX);
   END_IF;
END_REGION

REGION Network 87: R15 AUTO/MANUAL OUTPUT
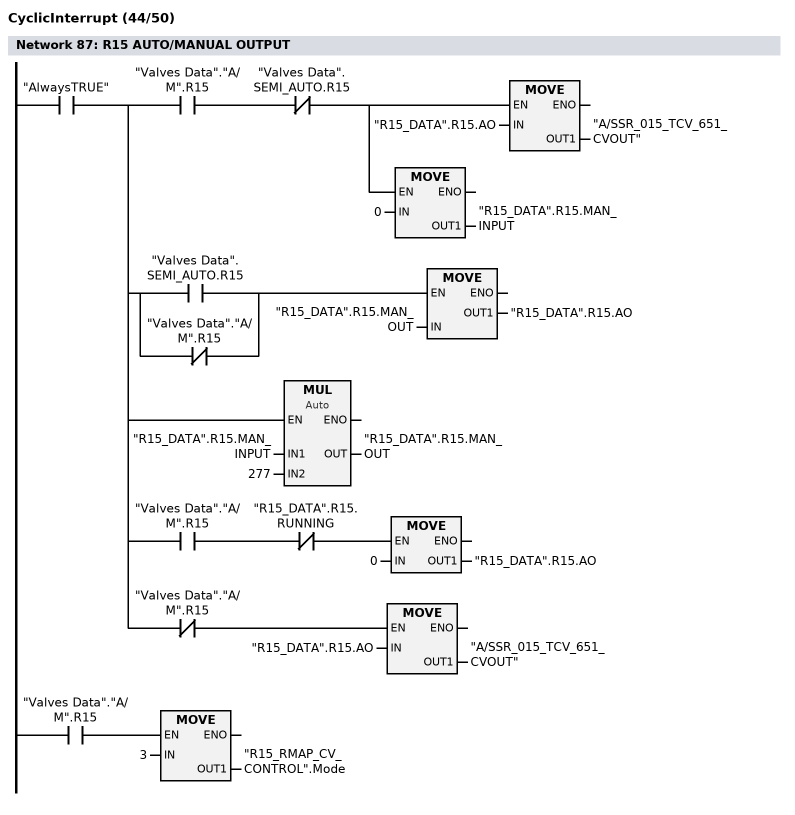
   RUNG wire#powerrail
      Contact( "AlwaysTRUE" )
      wire#w1
      Contact( "Valves Data"."A/M".R15 )
      I_Contact( "Valves Data".SEMI_AUTO.R15 )
      wire#w2
      Move(in := "R15_DATA".R15.AO, out1 => "A/SSR_015_TCV_651_CVOUT")
   END_RUNG
   RUNG wire#w2
      Move(in := 0, out1 => "R15_DATA".R15.MAN_INPUT)
   END_RUNG
   RUNG wire#w1
      Contact( "Valves Data".SEMI_AUTO.R15 )
      wire#w3
      Move(in := "R15_DATA".R15.MAN_OUT, out1 => "R15_DATA".R15.AO)
   END_RUNG
   RUNG wire#w1
      I_Contact( "Valves Data"."A/M".R15 )
   END_RUNG wire#w3
   RUNG wire#w1
      Mul(in1 := "R15_DATA".R15.MAN_INPUT, in2 := 277, out => "R15_DATA".R15.MAN_OUT)
   END_RUNG
   RUNG wire#w1
      Contact( "Valves Data"."A/M".R15 )
      I_Contact( "R15_DATA".R15.RUNNING )
      Move(in := 0, out1 => "R15_DATA".R15.AO)
   END_RUNG
   RUNG wire#w1
      I_Contact( "Valves Data"."A/M".R15 )
      Move(in := "R15_DATA".R15.AO, out1 => "A/SSR_015_TCV_651_CVOUT")
   END_RUNG
   RUNG wire#powerrail
      Contact( "Valves Data"."A/M".R15 )
      Move(in := 3, out1 => "R15_RMAP_CV_CONTROL".Mode)
   END_RUNG
   // the same network as SCL:
   IF "AlwaysTRUE" AND "Valves Data"."A/M".R15 AND NOT "Valves Data".SEMI_AUTO.R15 THEN
       "A/SSR_015_TCV_651_CVOUT" := "R15_DATA".R15.AO;
       "R15_DATA".R15.MAN_INPUT := 0;
   END_IF;
   IF "AlwaysTRUE" AND ("Valves Data".SEMI_AUTO.R15 OR NOT "Valves Data"."A/M".R15) THEN
       "R15_DATA".R15.AO := "R15_DATA".R15.MAN_OUT;
   END_IF;
   IF "AlwaysTRUE" THEN "R15_DATA".R15.MAN_OUT := "R15_DATA".R15.MAN_INPUT * 277; END_IF;
   IF "AlwaysTRUE" AND "Valves Data"."A/M".R15 AND NOT "R15_DATA".R15.RUNNING THEN
       "R15_DATA".R15.AO := 0;
   END_IF;
   IF "AlwaysTRUE" AND NOT "Valves Data"."A/M".R15 THEN
       "A/SSR_015_TCV_651_CVOUT" := "R15_DATA".R15.AO;
   END_IF;
   IF "Valves Data"."A/M".R15 THEN "R15_RMAP_CV_CONTROL".Mode := 3; END_IF;
END_REGION

REGION Network 88: R16_RAMP_CV
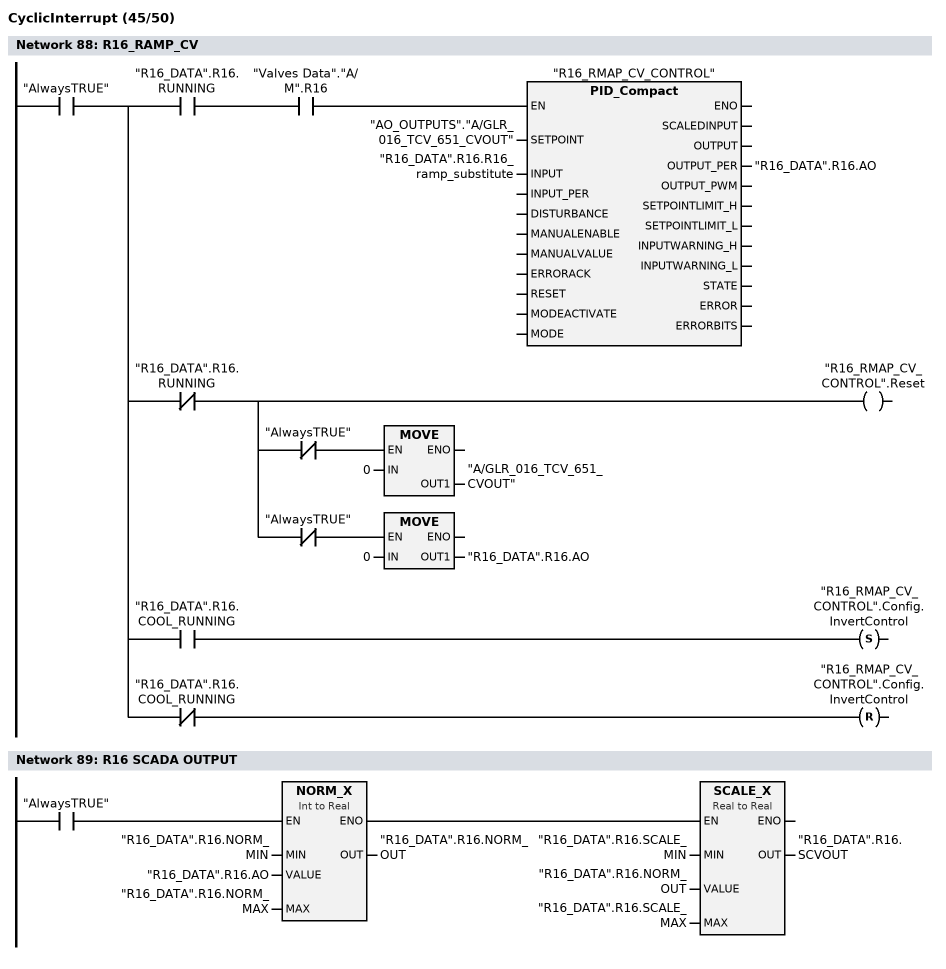
   RUNG wire#powerrail
      Contact( "AlwaysTRUE" )
      wire#w1
      Contact( "R16_DATA".R16.RUNNING )
      Contact( "Valves Data"."A/M".R16 )
      "R16_RMAP_CV_CONTROL".PID_Compact(Setpoint := "AO_OUTPUTS"."A/GLR_016_TCV_651_CVOUT", Input := "R16_DATA".R16.R16_ramp_substitute, Input_PER :=, Disturbance :=, ManualEnable :=, ManualValue :=, ErrorAck :=, Reset :=, ModeActivate :=, Mode :=, ScaledInput =>, Output =>, Output_PER => "R16_DATA".R16.AO, Output_PWM =>, SetpointLimit_H =>, SetpointLimit_L =>, InputWarning_H =>, InputWarning_L =>, State =>, Error =>, ErrorBits =>)
   END_RUNG
   RUNG wire#w1
      I_Contact( "R16_DATA".R16.RUNNING )
      wire#w2
      Coil( "R16_RMAP_CV_CONTROL".Reset )
   END_RUNG
   RUNG wire#w2
      I_Contact( "AlwaysTRUE" )
      Move(in := 0, out1 => "A/GLR_016_TCV_651_CVOUT")
   END_RUNG
   RUNG wire#w2
      I_Contact( "AlwaysTRUE" )
      Move(in := 0, out1 => "R16_DATA".R16.AO)
   END_RUNG
   RUNG wire#w1
      Contact( "R16_DATA".R16.COOL_RUNNING )
      S_Coil( "R16_RMAP_CV_CONTROL".Config.InvertControl )
   END_RUNG
   RUNG wire#w1
      I_Contact( "R16_DATA".R16.COOL_RUNNING )
      R_Coil( "R16_RMAP_CV_CONTROL".Config.InvertControl )
   END_RUNG
   // the same network as SCL:
   #_w1 := "AlwaysTRUE";
   IF "AlwaysTRUE" AND "R16_DATA".R16.RUNNING AND "Valves Data"."A/M".R16 THEN
       "R16_RMAP_CV_CONTROL"(Setpoint := "AO_OUTPUTS"."A/GLR_016_TCV_651_CVOUT",   // PID_Compact
                             Input := "R16_DATA".R16.R16_ramp_substitute,
                             Output_PER => "R16_DATA".R16.AO);
   END_IF;
   "R16_RMAP_CV_CONTROL".Reset := #_w1 AND NOT "R16_DATA".R16.RUNNING;
   IF "R16_RMAP_CV_CONTROL".Reset AND NOT "AlwaysTRUE" THEN
       "A/GLR_016_TCV_651_CVOUT" := 0;
       "R16_DATA".R16.AO := 0;
   END_IF;
   IF #_w1 AND "R16_DATA".R16.COOL_RUNNING THEN "R16_RMAP_CV_CONTROL".Config.InvertControl := TRUE; END_IF;
   IF #_w1 AND NOT "R16_DATA".R16.COOL_RUNNING THEN
       "R16_RMAP_CV_CONTROL".Config.InvertControl := FALSE;
   END_IF;
END_REGION

REGION Network 89: R16 SCADA OUTPUT
   RUNG wire#powerrail
      Contact( "AlwaysTRUE" )
      { S7_Templates := "[SrcType := Int, DestType := Real]" } Normalize(min := "R16_DATA".R16.NORM_MIN, value := "R16_DATA".R16.AO, max := "R16_DATA".R16.NORM_MAX, out => "R16_DATA".R16.NORM_OUT)
      { S7_Templates := "[SrcType := Real, DestType := Real]" } Scale(min := "R16_DATA".R16.SCALE_MIN, value := "R16_DATA".R16.NORM_OUT, max := "R16_DATA".R16.SCALE_MAX, out => "R16_DATA".R16.SCVOUT)
   END_RUNG
   // the same network as SCL:
   IF "AlwaysTRUE" THEN
       "R16_DATA".R16.NORM_OUT := NORM_X(MIN := "R16_DATA".R16.NORM_MIN, VALUE := "R16_DATA".R16.AO, MAX := "R16_DATA".R16.NORM_MAX);
       "R16_DATA".R16.SCVOUT := SCALE_X(MIN := "R16_DATA".R16.SCALE_MIN, VALUE := "R16_DATA".R16.NORM_OUT, MAX := "R16_DATA".R16.SCALE_MAX);
   END_IF;
END_REGION

REGION Network 90: R16 AUTO/MANUAL OUTPUT
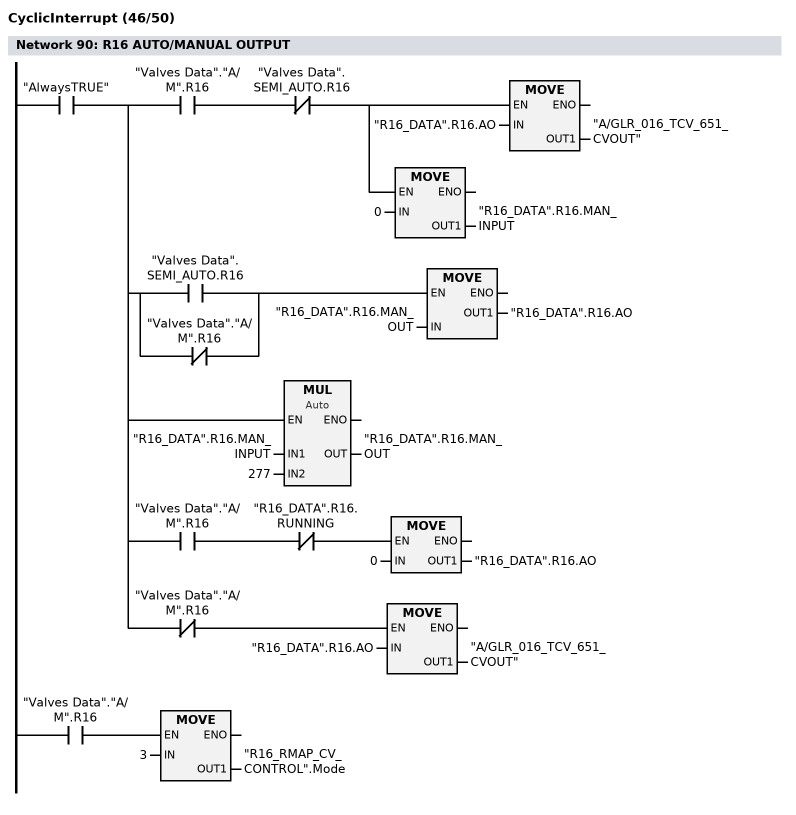
   RUNG wire#powerrail
      Contact( "AlwaysTRUE" )
      wire#w1
      Contact( "Valves Data"."A/M".R16 )
      I_Contact( "Valves Data".SEMI_AUTO.R16 )
      wire#w2
      Move(in := "R16_DATA".R16.AO, out1 => "A/GLR_016_TCV_651_CVOUT")
   END_RUNG
   RUNG wire#w2
      Move(in := 0, out1 => "R16_DATA".R16.MAN_INPUT)
   END_RUNG
   RUNG wire#w1
      Contact( "Valves Data".SEMI_AUTO.R16 )
      wire#w3
      Move(in := "R16_DATA".R16.MAN_OUT, out1 => "R16_DATA".R16.AO)
   END_RUNG
   RUNG wire#w1
      I_Contact( "Valves Data"."A/M".R16 )
   END_RUNG wire#w3
   RUNG wire#w1
      Mul(in1 := "R16_DATA".R16.MAN_INPUT, in2 := 277, out => "R16_DATA".R16.MAN_OUT)
   END_RUNG
   RUNG wire#w1
      Contact( "Valves Data"."A/M".R16 )
      I_Contact( "R16_DATA".R16.RUNNING )
      Move(in := 0, out1 => "R16_DATA".R16.AO)
   END_RUNG
   RUNG wire#w1
      I_Contact( "Valves Data"."A/M".R16 )
      Move(in := "R16_DATA".R16.AO, out1 => "A/GLR_016_TCV_651_CVOUT")
   END_RUNG
   RUNG wire#powerrail
      Contact( "Valves Data"."A/M".R16 )
      Move(in := 3, out1 => "R16_RMAP_CV_CONTROL".Mode)
   END_RUNG
   // the same network as SCL:
   IF "AlwaysTRUE" AND "Valves Data"."A/M".R16 AND NOT "Valves Data".SEMI_AUTO.R16 THEN
       "A/GLR_016_TCV_651_CVOUT" := "R16_DATA".R16.AO;
       "R16_DATA".R16.MAN_INPUT := 0;
   END_IF;
   IF "AlwaysTRUE" AND ("Valves Data".SEMI_AUTO.R16 OR NOT "Valves Data"."A/M".R16) THEN
       "R16_DATA".R16.AO := "R16_DATA".R16.MAN_OUT;
   END_IF;
   IF "AlwaysTRUE" THEN "R16_DATA".R16.MAN_OUT := "R16_DATA".R16.MAN_INPUT * 277; END_IF;
   IF "AlwaysTRUE" AND "Valves Data"."A/M".R16 AND NOT "R16_DATA".R16.RUNNING THEN
       "R16_DATA".R16.AO := 0;
   END_IF;
   IF "AlwaysTRUE" AND NOT "Valves Data"."A/M".R16 THEN
       "A/GLR_016_TCV_651_CVOUT" := "R16_DATA".R16.AO;
   END_IF;
   IF "Valves Data"."A/M".R16 THEN "R16_RMAP_CV_CONTROL".Mode := 3; END_IF;
END_REGION

REGION Network 91: R17_RAMP_CV
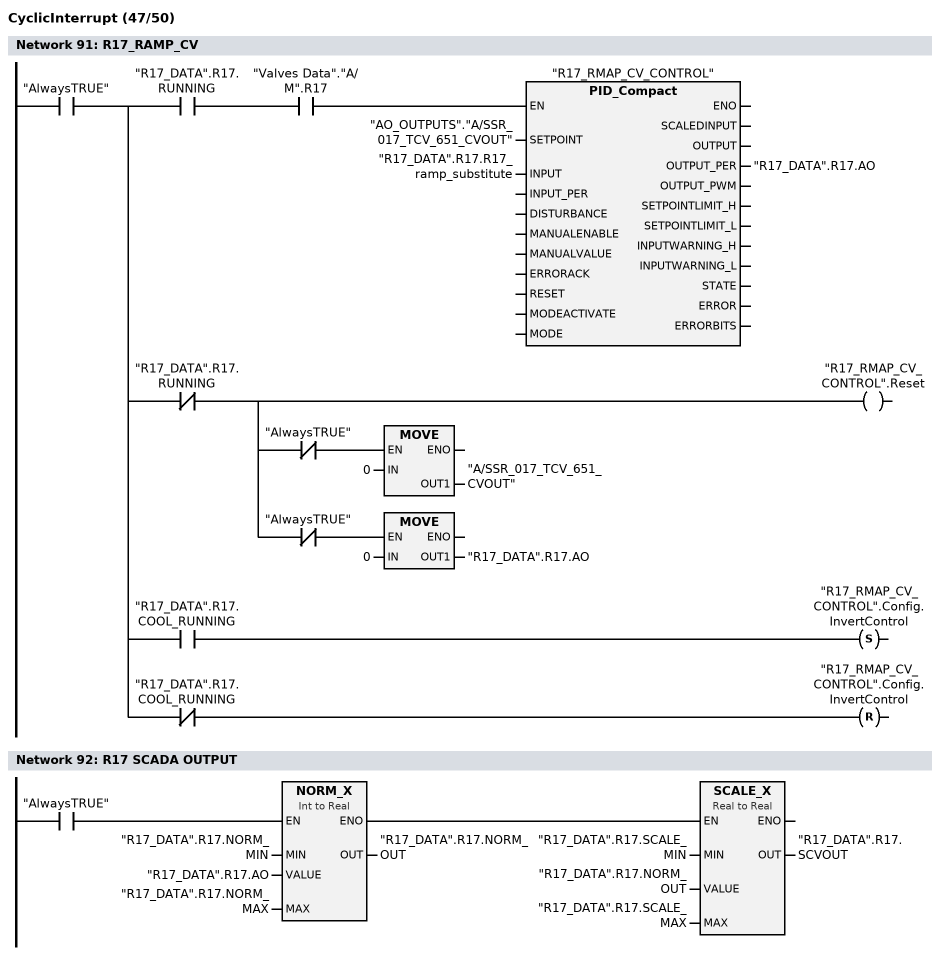
   RUNG wire#powerrail
      Contact( "AlwaysTRUE" )
      wire#w1
      Contact( "R17_DATA".R17.RUNNING )
      Contact( "Valves Data"."A/M".R17 )
      "R17_RMAP_CV_CONTROL".PID_Compact(Setpoint := "AO_OUTPUTS"."A/SSR_017_TCV_651_CVOUT", Input := "R17_DATA".R17.R17_ramp_substitute, Input_PER :=, Disturbance :=, ManualEnable :=, ManualValue :=, ErrorAck :=, Reset :=, ModeActivate :=, Mode :=, ScaledInput =>, Output =>, Output_PER => "R17_DATA".R17.AO, Output_PWM =>, SetpointLimit_H =>, SetpointLimit_L =>, InputWarning_H =>, InputWarning_L =>, State =>, Error =>, ErrorBits =>)
   END_RUNG
   RUNG wire#w1
      I_Contact( "R17_DATA".R17.RUNNING )
      wire#w2
      Coil( "R17_RMAP_CV_CONTROL".Reset )
   END_RUNG
   RUNG wire#w2
      I_Contact( "AlwaysTRUE" )
      Move(in := 0, out1 => "A/SSR_017_TCV_651_CVOUT")
   END_RUNG
   RUNG wire#w2
      I_Contact( "AlwaysTRUE" )
      Move(in := 0, out1 => "R17_DATA".R17.AO)
   END_RUNG
   RUNG wire#w1
      Contact( "R17_DATA".R17.COOL_RUNNING )
      S_Coil( "R17_RMAP_CV_CONTROL".Config.InvertControl )
   END_RUNG
   RUNG wire#w1
      I_Contact( "R17_DATA".R17.COOL_RUNNING )
      R_Coil( "R17_RMAP_CV_CONTROL".Config.InvertControl )
   END_RUNG
   // the same network as SCL:
   #_w1 := "AlwaysTRUE";
   IF "AlwaysTRUE" AND "R17_DATA".R17.RUNNING AND "Valves Data"."A/M".R17 THEN
       "R17_RMAP_CV_CONTROL"(Setpoint := "AO_OUTPUTS"."A/SSR_017_TCV_651_CVOUT",   // PID_Compact
                             Input := "R17_DATA".R17.R17_ramp_substitute,
                             Output_PER => "R17_DATA".R17.AO);
   END_IF;
   "R17_RMAP_CV_CONTROL".Reset := #_w1 AND NOT "R17_DATA".R17.RUNNING;
   IF "R17_RMAP_CV_CONTROL".Reset AND NOT "AlwaysTRUE" THEN
       "A/SSR_017_TCV_651_CVOUT" := 0;
       "R17_DATA".R17.AO := 0;
   END_IF;
   IF #_w1 AND "R17_DATA".R17.COOL_RUNNING THEN "R17_RMAP_CV_CONTROL".Config.InvertControl := TRUE; END_IF;
   IF #_w1 AND NOT "R17_DATA".R17.COOL_RUNNING THEN
       "R17_RMAP_CV_CONTROL".Config.InvertControl := FALSE;
   END_IF;
END_REGION

REGION Network 92: R17 SCADA OUTPUT
   RUNG wire#powerrail
      Contact( "AlwaysTRUE" )
      { S7_Templates := "[SrcType := Int, DestType := Real]" } Normalize(min := "R17_DATA".R17.NORM_MIN, value := "R17_DATA".R17.AO, max := "R17_DATA".R17.NORM_MAX, out => "R17_DATA".R17.NORM_OUT)
      { S7_Templates := "[SrcType := Real, DestType := Real]" } Scale(min := "R17_DATA".R17.SCALE_MIN, value := "R17_DATA".R17.NORM_OUT, max := "R17_DATA".R17.SCALE_MAX, out => "R17_DATA".R17.SCVOUT)
   END_RUNG
   // the same network as SCL:
   IF "AlwaysTRUE" THEN
       "R17_DATA".R17.NORM_OUT := NORM_X(MIN := "R17_DATA".R17.NORM_MIN, VALUE := "R17_DATA".R17.AO, MAX := "R17_DATA".R17.NORM_MAX);
       "R17_DATA".R17.SCVOUT := SCALE_X(MIN := "R17_DATA".R17.SCALE_MIN, VALUE := "R17_DATA".R17.NORM_OUT, MAX := "R17_DATA".R17.SCALE_MAX);
   END_IF;
END_REGION

REGION Network 93: R17 AUTO/MANUAL OUTPUT
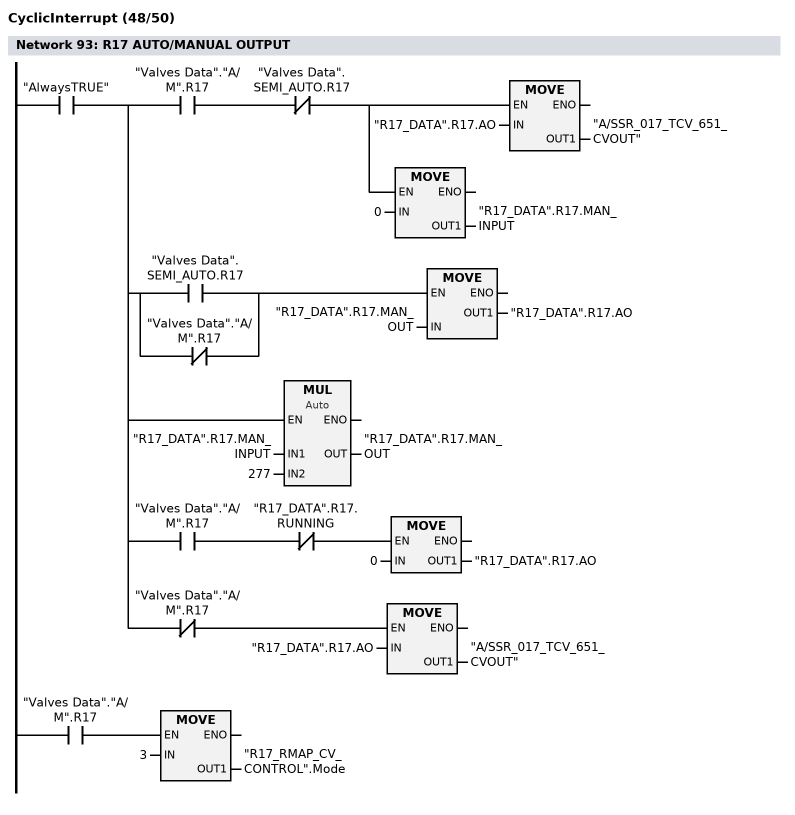
   RUNG wire#powerrail
      Contact( "AlwaysTRUE" )
      wire#w1
      Contact( "Valves Data"."A/M".R17 )
      I_Contact( "Valves Data".SEMI_AUTO.R17 )
      wire#w2
      Move(in := "R17_DATA".R17.AO, out1 => "A/SSR_017_TCV_651_CVOUT")
   END_RUNG
   RUNG wire#w2
      Move(in := 0, out1 => "R17_DATA".R17.MAN_INPUT)
   END_RUNG
   RUNG wire#w1
      Contact( "Valves Data".SEMI_AUTO.R17 )
      wire#w3
      Move(in := "R17_DATA".R17.MAN_OUT, out1 => "R17_DATA".R17.AO)
   END_RUNG
   RUNG wire#w1
      I_Contact( "Valves Data"."A/M".R17 )
   END_RUNG wire#w3
   RUNG wire#w1
      Mul(in1 := "R17_DATA".R17.MAN_INPUT, in2 := 277, out => "R17_DATA".R17.MAN_OUT)
   END_RUNG
   RUNG wire#w1
      Contact( "Valves Data"."A/M".R17 )
      I_Contact( "R17_DATA".R17.RUNNING )
      Move(in := 0, out1 => "R17_DATA".R17.AO)
   END_RUNG
   RUNG wire#w1
      I_Contact( "Valves Data"."A/M".R17 )
      Move(in := "R17_DATA".R17.AO, out1 => "A/SSR_017_TCV_651_CVOUT")
   END_RUNG
   RUNG wire#powerrail
      Contact( "Valves Data"."A/M".R17 )
      Move(in := 3, out1 => "R17_RMAP_CV_CONTROL".Mode)
   END_RUNG
   // the same network as SCL:
   IF "AlwaysTRUE" AND "Valves Data"."A/M".R17 AND NOT "Valves Data".SEMI_AUTO.R17 THEN
       "A/SSR_017_TCV_651_CVOUT" := "R17_DATA".R17.AO;
       "R17_DATA".R17.MAN_INPUT := 0;
   END_IF;
   IF "AlwaysTRUE" AND ("Valves Data".SEMI_AUTO.R17 OR NOT "Valves Data"."A/M".R17) THEN
       "R17_DATA".R17.AO := "R17_DATA".R17.MAN_OUT;
   END_IF;
   IF "AlwaysTRUE" THEN "R17_DATA".R17.MAN_OUT := "R17_DATA".R17.MAN_INPUT * 277; END_IF;
   IF "AlwaysTRUE" AND "Valves Data"."A/M".R17 AND NOT "R17_DATA".R17.RUNNING THEN
       "R17_DATA".R17.AO := 0;
   END_IF;
   IF "AlwaysTRUE" AND NOT "Valves Data"."A/M".R17 THEN
       "A/SSR_017_TCV_651_CVOUT" := "R17_DATA".R17.AO;
   END_IF;
   IF "Valves Data"."A/M".R17 THEN "R17_RMAP_CV_CONTROL".Mode := 3; END_IF;
END_REGION

REGION Network 94: R18_RAMP_CV
